--- program platizq (robot Fanuc LR Mate 200iD/7L) ---
  Suave(1)
  Establecer velocidad (1000.0 mm/s)
  Est. Ref.: RobotiQ 2F-140 Gripper (Mechanism) Base
  Est. herr: Tool 1
  Mostrar Tool 1
  MoveJ 1 to (260.93, 112.74, 317.18) mm, rotated rx -163.75 ry -45.95 rz -164.16 deg; joints [66.37, 34.682, -17.427, -50.975, -57.423, 69.366]
  MoveL 2 to (260.93, 112.74, 317.18) mm, rotated rx -163.75 ry -45.95 rz -164.16 deg; joints [66.37, 34.682, -17.427, -50.975, -57.423, 69.366]
  MoveL 3 to (241.32, 112.74, 219.12) mm, rotated rx -163.75 ry -45.95 rz -164.16 deg; joints [66.988, 41.165, -27.056, -56.554, -51.255, 78.508]
  MoveL 4 to (241.32, 112.74, 219.12) mm, rotated rx -163.75 ry -45.95 rz -164.16 deg; joints [66.988, 41.165, -27.056, -56.554, -51.255, 78.508]
  Establecer velocidad (50.0 mm/s)
  MoveL 5 to (253.05, 113.72, 219.12) mm, rotated rx -163.75 ry -45.95 rz -164.16 deg; joints [66.551, 39.855, -28.019, -57.172, -51.053, 79.816]
  MoveL 6 to (264.85, 113.71, 219.12) mm, rotated rx -163.75 ry -45.95 rz -164.16 deg; joints [66.172, 38.517, -28.983, -57.797, -50.815, 81.094]
  MoveL 7 to (276.61, 112.7, 219.12) mm, rotated rx -163.75 ry -45.95 rz -164.16 deg; joints [65.858, 37.162, -29.939, -58.425, -50.543, 82.329]
  MoveL 8 to (288.2, 110.7, 219.12) mm, rotated rx -163.75 ry -45.95 rz -164.16 deg; joints [65.614, 35.801, -30.876, -59.055, -50.236, 83.51]
  MoveL 9 to (299.55, 107.74, 219.66) mm, rotated rx -163.75 ry -45.95 rz -164.16 deg; joints [65.446, 34.407, -31.728, -59.642, -49.925, 84.562]
  MoveL 10 to (311.25, 103.8, 221.33) mm, rotated rx -163.75 ry -45.95 rz -164.16 deg; joints [65.334, 32.878, -32.469, -60.165, -49.635, 85.463]
  MoveL 11 to (322.85, 100.34, 224.12) mm, rotated rx -163.75 ry -45.95 rz -164.16 deg; joints [65.186, 31.325, -33.014, -60.541, -49.474, 86.167]
  MoveL 12 to (334.34, 97.51, 228.04) mm, rotated rx -163.75 ry -45.95 rz -164.16 deg; joints [64.983, 29.751, -33.357, -60.757, -49.454, 86.67]
  MoveL 13 to (346, 95.24, 231.53) mm, rotated rx -163.75 ry -45.95 rz -164.16 deg; joints [64.72, 28.217, -33.701, -60.96, -49.478, 87.205]
  MoveL 14 to (357.95, 93.53, 233.87) mm, rotated rx -163.75 ry -45.95 rz -164.16 deg; joints [64.39, 26.758, -34.143, -61.22, -49.504, 87.889]
  MoveL 15 to (370.19, 92.4, 235.02) mm, rotated rx -163.75 ry -45.95 rz -164.16 deg; joints [63.985, 25.377, -34.691, -61.538, -49.535, 88.731]
  MoveL 16 to (383.51, 91.88, 235.15) mm, rotated rx -163.75 ry -45.95 rz -164.16 deg; joints [63.465, 23.993, -35.369, -61.92, -49.589, 89.781]
  MoveL 17 to (396.84, 92.08, 235.15) mm, rotated rx -163.75 ry -45.95 rz -164.16 deg; joints [62.858, 22.663, -36.01, -62.244, -49.724, 90.827]
  MoveL 18 to (410.17, 92.08, 235.15) mm, rotated rx -163.75 ry -45.95 rz -164.16 deg; joints [62.245, 21.332, -36.621, -62.531, -49.879, 91.835]
  MoveL 19 to (423.5, 92.08, 235.15) mm, rotated rx -163.75 ry -45.95 rz -164.16 deg; joints [61.606, 20.009, -37.197, -62.774, -50.068, 92.81]
  MoveL 20 to (436.83, 92.08, 235.15) mm, rotated rx -163.75 ry -45.95 rz -164.16 deg; joints [60.939, 18.692, -37.738, -62.971, -50.292, 93.751]
  MoveL 21 to (445.16, 92.08, 235.15) mm, rotated rx -163.75 ry -45.95 rz -164.16 deg; joints [60.508, 17.872, -38.059, -63.071, -50.45, 94.323]
  MoveL 22 to (453.49, 92.08, 235.15) mm, rotated rx -163.75 ry -45.95 rz -164.16 deg; joints [60.065, 17.054, -38.366, -63.152, -50.622, 94.881]
  MoveL 23 to (461.82, 92.08, 235.15) mm, rotated rx -163.75 ry -45.95 rz -164.16 deg; joints [59.609, 16.238, -38.659, -63.214, -50.808, 95.427]
  MoveL 24 to (470.22, 91.84, 235.15) mm, rotated rx -163.75 ry -45.95 rz -164.16 deg; joints [59.16, 15.403, -38.947, -63.269, -50.991, 95.961]
  MoveL 25 to (476.05, 90.4, 235.15) mm, rotated rx -163.75 ry -45.95 rz -164.16 deg; joints [58.963, 14.749, -39.161, -63.356, -51.031, 96.296]
  MoveL 26 to (481.67, 87.57, 235.15) mm, rotated rx -163.75 ry -45.95 rz -164.16 deg; joints [58.91, 14.031, -39.387, -63.501, -50.967, 96.58]
  MoveL 27 to (486.6, 83.43, 235.15) mm, rotated rx -163.75 ry -45.95 rz -164.16 deg; joints [59.025, 13.302, -39.606, -63.701, -50.79, 96.782]
  MoveL 28 to (490.42, 78.28, 235.15) mm, rotated rx -163.75 ry -45.95 rz -164.16 deg; joints [59.311, 12.621, -39.801, -63.948, -50.507, 96.882]
  MoveL 29 to (492.88, 72.58, 235.15) mm, rotated rx -163.75 ry -45.95 rz -164.16 deg; joints [59.741, 12.041, -39.958, -64.221, -50.141, 96.879]
  MoveL 30 to (493.98, 66.8, 235.15) mm, rotated rx -163.75 ry -45.95 rz -164.16 deg; joints [60.268, 11.597, -40.075, -64.502, -49.727, 96.788]
  MoveL 31 to (494.07, 61.23, 235.15) mm, rotated rx -163.75 ry -45.95 rz -164.16 deg; joints [60.841, 11.27, -40.158, -64.774, -49.296, 96.64]
  MoveL 32 to (494.07, 55.68, 235.15) mm, rotated rx -163.75 ry -45.95 rz -164.16 deg; joints [61.423, 10.958, -40.235, -65.047, -48.86, 96.482]
  MoveL 33 to (493.53, 50, 235.15) mm, rotated rx -163.75 ry -45.95 rz -164.16 deg; joints [62.056, 10.7, -40.297, -65.328, -48.395, 96.287]
  MoveL 34 to (491.67, 44.21, 235.15) mm, rotated rx -163.75 ry -45.95 rz -164.16 deg; joints [62.78, 10.579, -40.325, -65.614, -47.881, 96.014]
  MoveL 35 to (488.43, 38.76, 235.15) mm, rotated rx -163.75 ry -45.95 rz -164.16 deg; joints [63.546, 10.629, -40.313, -65.88, -47.354, 95.675]
  MoveL 36 to (483.95, 34.13, 235.15) mm, rotated rx -163.75 ry -45.95 rz -164.16 deg; joints [64.285, 10.862, -40.258, -66.098, -46.861, 95.292]
  MoveL 37 to (478.57, 30.7, 235.15) mm, rotated rx -163.75 ry -45.95 rz -164.16 deg; joints [64.933, 11.256, -40.161, -66.244, -46.448, 94.895]
  MoveL 38 to (472.77, 28.65, 235.15) mm, rotated rx -163.75 ry -45.95 rz -164.16 deg; joints [65.443, 11.768, -40.03, -66.308, -46.143, 94.513]
  MoveL 39 to (465.18, 27.94, 235.15) mm, rotated rx -163.75 ry -45.95 rz -164.16 deg; joints [65.887, 12.534, -39.824, -66.279, -45.915, 94.061]
  MoveL 40 to (457.78, 27.94, 235.15) mm, rotated rx -163.75 ry -45.95 rz -164.16 deg; joints [66.235, 13.314, -39.602, -66.199, -45.759, 93.627]
  MoveL 41 to (450.37, 27.94, 235.15) mm, rotated rx -163.75 ry -45.95 rz -164.16 deg; joints [66.574, 14.092, -39.368, -66.103, -45.614, 93.18]
  MoveL 42 to (442.97, 27.94, 235.15) mm, rotated rx -163.75 ry -45.95 rz -164.16 deg; joints [66.905, 14.869, -39.122, -65.989, -45.48, 92.719]
  MoveL 43 to (435.56, 27.94, 235.15) mm, rotated rx -163.75 ry -45.95 rz -164.16 deg; joints [67.226, 15.646, -38.864, -65.859, -45.357, 92.245]
  MoveL 44 to (428.16, 27.94, 235.15) mm, rotated rx -163.75 ry -45.95 rz -164.16 deg; joints [67.539, 16.422, -38.594, -65.712, -45.245, 91.758]
  MoveL 45 to (413.49, 27.94, 235.15) mm, rotated rx -163.75 ry -45.95 rz -164.16 deg; joints [68.135, 17.958, -38.025, -65.374, -45.055, 90.755]
  MoveL 46 to (398.83, 27.94, 235.15) mm, rotated rx -163.75 ry -45.95 rz -164.16 deg; joints [68.702, 19.495, -37.412, -64.975, -44.906, 89.701]
  MoveL 47 to (384.18, 27.45, 235.15) mm, rotated rx -163.75 ry -45.95 rz -164.16 deg; joints [69.288, 21.014, -36.762, -64.536, -44.76, 88.584]
  MoveL 48 to (369.59, 25.97, 235) mm, rotated rx -163.75 ry -45.95 rz -164.16 deg; joints [69.936, 22.505, -36.108, -64.097, -44.573, 87.425]
  MoveL 49 to (357.46, 23.95, 233.79) mm, rotated rx -163.75 ry -45.95 rz -164.16 deg; joints [70.525, 23.796, -35.681, -63.837, -44.332, 86.577]
  MoveL 50 to (345.61, 21.29, 231.44) mm, rotated rx -163.75 ry -45.95 rz -164.16 deg; joints [71.143, 25.115, -35.39, -63.699, -44.01, 85.885]
  MoveL 51 to (334.07, 18.15, 227.95) mm, rotated rx -163.75 ry -45.95 rz -164.16 deg; joints [71.773, 26.466, -35.228, -63.675, -43.621, 85.346]
  MoveL 52 to (322.58, 15.47, 224.04) mm, rotated rx -163.75 ry -45.95 rz -164.16 deg; joints [72.34, 27.861, -35.073, -63.637, -43.274, 84.844]
  MoveL 53 to (310.79, 13.36, 221.24) mm, rotated rx -163.75 ry -45.95 rz -164.16 deg; joints [72.848, 29.241, -34.718, -63.39, -43.059, 84.107]
  MoveL 54 to (298.7, 11.85, 219.58) mm, rotated rx -163.75 ry -45.95 rz -164.16 deg; joints [73.295, 30.606, -34.158, -62.93, -42.983, 83.131]
  MoveL 55 to (287.65, 11.04, 219.12) mm, rotated rx -163.75 ry -45.95 rz -164.16 deg; joints [73.643, 31.816, -33.482, -62.337, -43.037, 82.057]
  MoveL 56 to (276.52, 10.76, 219.12) mm, rotated rx -163.75 ry -45.95 rz -164.16 deg; joints [73.937, 33.036, -32.706, -61.643, -43.184, 80.886]
  MoveL 57 to (265.38, 10.76, 219.12) mm, rotated rx -163.75 ry -45.95 rz -164.16 deg; joints [74.199, 34.28, -31.895, -60.914, -43.38, 79.692]
  MoveL 58 to (254.26, 11.36, 219.12) mm, rotated rx -163.75 ry -45.95 rz -164.16 deg; joints [74.404, 35.558, -31.04, -60.146, -43.648, 78.486]
  MoveL 59 to (243.27, 13.24, 219.12) mm, rotated rx -163.75 ry -45.95 rz -164.16 deg; joints [74.498, 36.878, -30.135, -59.338, -44.034, 77.299]
  MoveL 60 to (232.6, 16.36, 219.32) mm, rotated rx -163.75 ry -45.95 rz -164.16 deg; joints [74.486, 38.214, -29.168, -58.488, -44.543, 76.121]
  MoveL 61 to (222.4, 20.67, 219.99) mm, rotated rx -163.75 ry -45.95 rz -164.16 deg; joints [74.372, 39.53, -28.125, -57.598, -45.18, 74.941]
  MoveL 62 to (212.73, 26.14, 221.07) mm, rotated rx -163.75 ry -45.95 rz -164.16 deg; joints [74.162, 40.83, -27.015, -56.685, -45.938, 73.777]
  MoveL 63 to (203.82, 32.62, 222.45) mm, rotated rx -163.75 ry -45.95 rz -164.16 deg; joints [73.867, 42.091, -25.876, -55.791, -46.791, 72.672]
  MoveL 64 to (198.88, 36.96, 223.38) mm, rotated rx -163.75 ry -45.95 rz -164.16 deg; joints [73.652, 42.825, -25.188, -55.273, -47.34, 72.046]
  MoveL 65 to (194.23, 41.63, 224.35) mm, rotated rx -163.75 ry -45.95 rz -164.16 deg; joints [73.409, 43.547, -24.498, -54.77, -47.917, 71.452]
  MoveL 66 to (189.92, 46.67, 225.35) mm, rotated rx -163.75 ry -45.95 rz -164.16 deg; joints [73.136, 44.252, -23.813, -54.289, -48.517, 70.898]
  MoveL 67 to (186.72, 52.48, 226.16) mm, rotated rx -163.75 ry -45.95 rz -164.16 deg; joints [72.787, 44.867, -23.221, -53.895, -49.123, 70.51]
  MoveL 68 to (185.04, 58.92, 226.6) mm, rotated rx -163.75 ry -45.95 rz -164.16 deg; joints [72.362, 45.336, -22.794, -53.631, -49.691, 70.36]
  MoveL 69 to (184.83, 66.37, 226.66) mm, rotated rx -163.75 ry -45.95 rz -164.16 deg; joints [71.836, 45.682, -22.514, -53.482, -50.247, 70.444]
  MoveL 70 to (185.41, 73.79, 226.5) mm, rotated rx -163.75 ry -45.95 rz -164.16 deg; joints [71.297, 45.942, -22.332, -53.401, -50.756, 70.64]
  MoveL 71 to (187.29, 80.95, 226.01) mm, rotated rx -163.75 ry -45.95 rz -164.16 deg; joints [70.746, 46.04, -22.325, -53.433, -51.17, 71.023]
  MoveL 72 to (190.4, 87.61, 225.24) mm, rotated rx -163.75 ry -45.95 rz -164.16 deg; joints [70.2, 45.976, -22.486, -53.568, -51.48, 71.573]
  MoveL 73 to (194.64, 93.62, 224.26) mm, rotated rx -163.75 ry -45.95 rz -164.16 deg; joints [69.67, 45.75, -22.802, -53.797, -51.687, 72.268]
  MoveL 74 to (199.85, 98.76, 223.19) mm, rotated rx -163.75 ry -45.95 rz -164.16 deg; joints [69.172, 45.372, -23.254, -54.102, -51.792, 73.077]
  MoveL 75 to (205.9, 102.91, 222.1) mm, rotated rx -163.75 ry -45.95 rz -164.16 deg; joints [68.717, 44.852, -23.817, -54.472, -51.802, 73.968]
  MoveL 76 to (212.58, 105.92, 221.09) mm, rotated rx -163.75 ry -45.95 rz -164.16 deg; joints [68.319, 44.205, -24.463, -54.89, -51.724, 74.907]
  MoveL 77 to (219.61, 108.2, 220.26) mm, rotated rx -163.75 ry -45.95 rz -164.16 deg; joints [67.958, 43.487, -25.137, -55.324, -51.608, 75.85]
  MoveL 78 to (226.74, 110.09, 219.65) mm, rotated rx -163.75 ry -45.95 rz -164.16 deg; joints [67.616, 42.741, -25.794, -55.746, -51.49, 76.765]
  MoveL 79 to (233.98, 111.61, 219.26) mm, rotated rx -163.75 ry -45.95 rz -164.16 deg; joints [67.293, 41.968, -26.434, -56.156, -51.373, 77.652]
  MoveL 80 to (241.32, 112.74, 219.12) mm, rotated rx -163.75 ry -45.95 rz -164.16 deg; joints [66.988, 41.165, -27.056, -56.554, -51.255, 78.508]
  Establecer velocidad (1000.0 mm/s)
  MoveL 81 to (241.32, 112.74, 219.12) mm, rotated rx -163.75 ry -45.95 rz -164.16 deg; joints [66.988, 41.165, -27.056, -56.554, -51.255, 78.508]
  MoveL 82 to (260.93, 112.74, 317.18) mm, rotated rx -163.75 ry -45.95 rz -164.16 deg; joints [66.37, 34.682, -17.427, -50.975, -57.423, 69.366]
  Establecer velocidad (1000.0 mm/s)
  MoveL 83 to (452.25, 27.76, 382.46) mm, rotated rx -163.75 ry -45.95 rz -164.16 deg; joints [66.508, 5.685, -18.926, -51.728, -56.385, 70.666]
  MoveL 84 to (432.64, 27.76, 284.4) mm, rotated rx -163.75 ry -45.95 rz -164.16 deg; joints [67.369, 12.539, -31.994, -60.148, -48.379, 83.782]
  MoveL 85 to (432.64, 27.76, 284.4) mm, rotated rx -163.75 ry -45.95 rz -164.16 deg; joints [67.369, 12.539, -31.994, -60.148, -48.379, 83.782]
  Establecer velocidad (50.0 mm/s)
  MoveL 86 to (452.8, 28.72, 284.4) mm, rotated rx -163.75 ry -45.95 rz -164.16 deg; joints [66.383, 10.356, -32.504, -60.376, -48.85, 84.924]
  MoveL 87 to (472.8, 31.52, 284.4) mm, rotated rx -163.75 ry -45.95 rz -164.16 deg; joints [65.133, 8.281, -32.901, -60.447, -49.569, 86.066]
  MoveL 88 to (479.3, 33.32, 284.4) mm, rotated rx -163.75 ry -45.95 rz -164.16 deg; joints [64.612, 7.655, -33.003, -60.422, -49.899, 86.466]
  MoveL 89 to (485.2, 36.51, 284.4) mm, rotated rx -163.75 ry -45.95 rz -164.16 deg; joints [63.96, 7.172, -33.077, -60.346, -50.337, 86.901]
  MoveL 90 to (490.31, 40.91, 284.4) mm, rotated rx -163.75 ry -45.95 rz -164.16 deg; joints [63.21, 6.849, -33.124, -60.226, -50.859, 87.357]
  MoveL 91 to (494.31, 46.34, 284.4) mm, rotated rx -163.75 ry -45.95 rz -164.16 deg; joints [62.404, 6.717, -33.143, -60.069, -51.436, 87.809]
  MoveL 92 to (496.77, 52.59, 284.4) mm, rotated rx -163.75 ry -45.95 rz -164.16 deg; joints [61.595, 6.811, -33.13, -59.885, -52.029, 88.226]
  MoveL 93 to (497.4, 59.25, 284.4) mm, rotated rx -163.75 ry -45.95 rz -164.16 deg; joints [60.853, 7.137, -33.083, -59.69, -52.589, 88.57]
  MoveL 94 to (497.21, 64.6, 284.4) mm, rotated rx -163.75 ry -45.95 rz -164.16 deg; joints [60.305, 7.479, -33.031, -59.534, -53.012, 88.806]
  MoveL 95 to (495.99, 69.73, 284.4) mm, rotated rx -163.75 ry -45.95 rz -164.16 deg; joints [59.846, 7.923, -32.961, -59.385, -53.379, 88.975]
  MoveL 96 to (493.74, 74.55, 284.4) mm, rotated rx -163.75 ry -45.95 rz -164.16 deg; joints [59.489, 8.458, -32.871, -59.247, -53.683, 89.068]
  MoveL 97 to (490.6, 78.79, 284.4) mm, rotated rx -163.75 ry -45.95 rz -164.16 deg; joints [59.249, 9.05, -32.764, -59.125, -53.911, 89.083]
  MoveL 98 to (486.76, 82.45, 284.4) mm, rotated rx -163.75 ry -45.95 rz -164.16 deg; joints [59.112, 9.678, -32.643, -59.019, -54.071, 89.028]
  MoveL 99 to (480.86, 86.17, 284.4) mm, rotated rx -163.75 ry -45.95 rz -164.16 deg; joints [59.093, 10.521, -32.469, -58.907, -54.175, 88.854]
  MoveL 100 to (474.22, 88.37, 284.4) mm, rotated rx -163.75 ry -45.95 rz -164.16 deg; joints [59.264, 11.343, -32.285, -58.831, -54.146, 88.568]
  MoveL 101 to (467.32, 89.52, 284.4) mm, rotated rx -163.75 ry -45.95 rz -164.16 deg; joints [59.546, 12.127, -32.098, -58.775, -54.04, 88.218]
  MoveL 102 to (460.39, 90.46, 284.4) mm, rotated rx -163.75 ry -45.95 rz -164.16 deg; joints [59.842, 12.9, -31.901, -58.715, -53.927, 87.849]
  MoveL 103 to (453.43, 91.18, 284.4) mm, rotated rx -163.75 ry -45.95 rz -164.16 deg; joints [60.152, 13.663, -31.696, -58.651, -53.808, 87.462]
  MoveL 104 to (446.45, 91.7, 284.4) mm, rotated rx -163.75 ry -45.95 rz -164.16 deg; joints [60.476, 14.416, -31.482, -58.581, -53.685, 87.058]
  MoveL 105 to (429.96, 92.12, 284.4) mm, rotated rx -163.75 ry -45.95 rz -164.16 deg; joints [61.282, 16.152, -30.948, -58.396, -53.375, 86.043]
  MoveL 106 to (413.48, 91.53, 284.4) mm, rotated rx -163.75 ry -45.95 rz -164.16 deg; joints [62.137, 17.84, -30.376, -58.179, -53.05, 84.952]
  MoveL 107 to (403.76, 90.49, 284.4) mm, rotated rx -163.75 ry -45.95 rz -164.16 deg; joints [62.684, 18.804, -30.026, -58.041, -52.834, 84.267]
  MoveL 108 to (394.19, 88.84, 284.4) mm, rotated rx -163.75 ry -45.95 rz -164.16 deg; joints [63.262, 19.726, -29.675, -57.9, -52.595, 83.559]
  MoveL 109 to (384.65, 87.33, 284.4) mm, rotated rx -163.75 ry -45.95 rz -164.16 deg; joints [63.811, 20.66, -29.304, -57.734, -52.389, 82.843]
  MoveL 110 to (374.95, 87.44, 284.4) mm, rotated rx -163.75 ry -45.95 rz -164.16 deg; joints [64.212, 21.702, -28.873, -57.503, -52.323, 82.146]
  MoveL 111 to (365.25, 87.59, 284.4) mm, rotated rx -163.75 ry -45.95 rz -164.16 deg; joints [64.598, 22.751, -28.42, -57.252, -52.282, 81.433]
  MoveL 112 to (355.55, 87.57, 284.4) mm, rotated rx -163.75 ry -45.95 rz -164.16 deg; joints [64.987, 23.799, -27.949, -56.986, -52.25, 80.697]
  MoveL 113 to (351.15, 87.43, 284.4) mm, rotated rx -163.75 ry -45.95 rz -164.16 deg; joints [65.171, 24.271, -27.731, -56.861, -52.233, 80.354]
  MoveL 114 to (346.75, 87.18, 284.4) mm, rotated rx -163.75 ry -45.95 rz -164.16 deg; joints [65.362, 24.738, -27.511, -56.736, -52.211, 80.004]
  MoveL 115 to (342.36, 86.74, 284.4) mm, rotated rx -163.75 ry -45.95 rz -164.16 deg; joints [65.565, 25.196, -27.293, -56.611, -52.181, 79.647]
  MoveL 116 to (338.08, 85.69, 284.4) mm, rotated rx -163.75 ry -45.95 rz -164.16 deg; joints [65.813, 25.614, -27.09, -56.498, -52.108, 79.28]
  MoveL 117 to (334.49, 83.14, 284.4) mm, rotated rx -163.75 ry -45.95 rz -164.16 deg; joints [66.158, 25.885, -26.957, -56.436, -51.926, 78.924]
  MoveL 118 to (332.28, 80.19, 284.4) mm, rotated rx -163.75 ry -45.95 rz -164.16 deg; joints [66.483, 25.986, -26.907, -56.424, -51.712, 78.667]
  MoveL 119 to (331.08, 76.71, 284.4) mm, rotated rx -163.75 ry -45.95 rz -164.16 deg; joints [66.815, 25.953, -26.924, -56.456, -51.456, 78.475]
  MoveL 120 to (331.16, 73.04, 284.4) mm, rotated rx -163.75 ry -45.95 rz -164.16 deg; joints [67.118, 25.771, -27.013, -56.534, -51.181, 78.38]
  MoveL 121 to (332.81, 67.76, 284.4) mm, rotated rx -163.75 ry -45.95 rz -164.16 deg; joints [67.503, 25.341, -27.222, -56.698, -50.78, 78.362]
  MoveL 122 to (334.61, 62.54, 284.4) mm, rotated rx -163.75 ry -45.95 rz -164.16 deg; joints [67.883, 24.902, -27.433, -56.865, -50.382, 78.351]
  MoveL 123 to (334.06, 60.19, 284.4) mm, rotated rx -163.75 ry -45.95 rz -164.16 deg; joints [68.102, 24.858, -27.454, -56.892, -50.208, 78.236]
  MoveL 124 to (333.37, 57.83, 284.4) mm, rotated rx -163.75 ry -45.95 rz -164.16 deg; joints [68.327, 24.83, -27.467, -56.914, -50.034, 78.109]
  MoveL 125 to (332.69, 55.47, 284.4) mm, rotated rx -163.75 ry -45.95 rz -164.16 deg; joints [68.552, 24.802, -27.481, -56.936, -49.859, 77.981]
  MoveL 126 to (332.02, 53.1, 284.4) mm, rotated rx -163.75 ry -45.95 rz -164.16 deg; joints [68.776, 24.773, -27.494, -56.957, -49.685, 77.853]
  MoveL 127 to (331.37, 50.73, 284.4) mm, rotated rx -163.75 ry -45.95 rz -164.16 deg; joints [69.001, 24.743, -27.508, -56.979, -49.51, 77.726]
  MoveL 128 to (330.99, 48.32, 284.4) mm, rotated rx -163.75 ry -45.95 rz -164.16 deg; joints [69.221, 24.682, -27.537, -57.01, -49.331, 77.618]
  MoveL 129 to (331.56, 43.51, 284.4) mm, rotated rx -163.75 ry -45.95 rz -164.16 deg; joints [69.618, 24.415, -27.663, -57.12, -48.967, 77.505]
  MoveL 130 to (333.68, 39.14, 284.4) mm, rotated rx -163.75 ry -45.95 rz -164.16 deg; joints [69.931, 23.996, -27.858, -57.278, -48.629, 77.523]
  MoveL 131 to (336.88, 35.49, 284.4) mm, rotated rx -163.75 ry -45.95 rz -164.16 deg; joints [70.148, 23.487, -28.091, -57.461, -48.342, 77.647]
  MoveL 132 to (341.1, 33.11, 284.4) mm, rotated rx -163.75 ry -45.95 rz -164.16 deg; joints [70.224, 22.917, -28.346, -57.658, -48.148, 77.888]
  MoveL 133 to (345.9, 32.32, 284.4) mm, rotated rx -163.75 ry -45.95 rz -164.16 deg; joints [70.141, 22.346, -28.597, -57.843, -48.076, 78.224]
  MoveL 134 to (350.74, 31.87, 284.4) mm, rotated rx -163.75 ry -45.95 rz -164.16 deg; joints [70.024, 21.785, -28.837, -58.019, -48.036, 78.572]
  MoveL 135 to (355.61, 31.66, 284.4) mm, rotated rx -163.75 ry -45.95 rz -164.16 deg; joints [69.883, 21.233, -29.069, -58.186, -48.018, 78.924]
  MoveL 136 to (360.47, 31.61, 284.4) mm, rotated rx -163.75 ry -45.95 rz -164.16 deg; joints [69.725, 20.689, -29.292, -58.346, -48.018, 79.277]
  MoveL 137 to (365.34, 31.66, 284.4) mm, rotated rx -163.75 ry -45.95 rz -164.16 deg; joints [69.554, 20.149, -29.508, -58.498, -48.031, 79.63]
  MoveL 138 to (370.79, 31.8, 284.4) mm, rotated rx -163.75 ry -45.95 rz -164.16 deg; joints [69.353, 19.55, -29.743, -58.66, -48.059, 80.021]
  MoveL 139 to (376.24, 31.99, 284.4) mm, rotated rx -163.75 ry -45.95 rz -164.16 deg; joints [69.144, 18.953, -29.969, -58.814, -48.096, 80.408]
  MoveL 140 to (381.69, 32.16, 284.4) mm, rotated rx -163.75 ry -45.95 rz -164.16 deg; joints [68.933, 18.357, -30.189, -58.962, -48.139, 80.788]
  MoveL 141 to (387.14, 32.28, 284.4) mm, rotated rx -163.75 ry -45.95 rz -164.16 deg; joints [68.722, 17.76, -30.404, -59.104, -48.184, 81.16]
  MoveL 142 to (392.5, 31.25, 284.4) mm, rotated rx -163.75 ry -45.95 rz -164.16 deg; joints [68.622, 17.124, -30.624, -59.262, -48.145, 81.474]
  MoveL 143 to (397.9, 29.94, 284.4) mm, rotated rx -163.75 ry -45.95 rz -164.16 deg; joints [68.544, 16.472, -30.844, -59.422, -48.091, 81.773]
  MoveL 144 to (403.83, 28.61, 284.4) mm, rotated rx -163.75 ry -45.95 rz -164.16 deg; joints [68.447, 15.758, -31.074, -59.589, -48.046, 82.097]
  MoveL 145 to (408.55, 28, 284.4) mm, rotated rx -163.75 ry -45.95 rz -164.16 deg; joints [68.324, 15.211, -31.244, -59.705, -48.051, 82.366]
  MoveL 146 to (412.24, 27.79, 284.4) mm, rotated rx -163.75 ry -45.95 rz -164.16 deg; joints [68.2, 14.793, -31.37, -59.786, -48.079, 82.584]
  MoveL 147 to (415.69, 27.76, 284.4) mm, rotated rx -163.75 ry -45.95 rz -164.16 deg; joints [68.066, 14.411, -31.483, -59.855, -48.121, 82.792]
  MoveL 148 to (418.69, 27.76, 284.4) mm, rotated rx -163.75 ry -45.95 rz -164.16 deg; joints [67.946, 14.08, -31.578, -59.912, -48.162, 82.971]
  MoveL 149 to (422.53, 27.76, 284.4) mm, rotated rx -163.75 ry -45.95 rz -164.16 deg; joints [67.79, 13.656, -31.697, -59.982, -48.217, 83.199]
  MoveL 150 to (427.35, 27.76, 284.4) mm, rotated rx -163.75 ry -45.95 rz -164.16 deg; joints [67.591, 13.123, -31.842, -60.064, -48.292, 83.48]
  MoveL 151 to (432.64, 27.76, 284.4) mm, rotated rx -163.75 ry -45.95 rz -164.16 deg; joints [67.369, 12.539, -31.994, -60.148, -48.379, 83.782]
  Establecer velocidad (1000.0 mm/s)
  MoveL 152 to (432.64, 27.76, 284.4) mm, rotated rx -163.75 ry -45.95 rz -164.16 deg; joints [67.369, 12.539, -31.994, -60.148, -48.379, 83.782]
  MoveL 153 to (452.25, 27.76, 382.46) mm, rotated rx -163.75 ry -45.95 rz -164.16 deg; joints [66.508, 5.685, -18.926, -51.728, -56.385, 70.666]

--- program carribizq (robot Fanuc LR Mate 200iD/7L) ---
  Suave(1)
  Establecer velocidad (1000.0 mm/s)
  Est. Ref.: RobotiQ 2F-140 Gripper (Mechanism) Base
  Est. herr: Tool 1
  Mostrar Tool 1
  MoveJ 1 to (259.22, -163.5, 158.15) mm, rotated rx 167 ry 29.36 rz -96.45 deg; joints [108.037, 52.448, -19.707, 33.515, -72.983, 58.084]
  MoveL 2 to (259.22, -163.5, 158.15) mm, rotated rx 167 ry 29.36 rz -96.45 deg; joints [108.037, 52.448, -19.707, 33.515, -72.983, 58.084]
  MoveL 3 to (239.61, -163.5, 60.09) mm, rotated rx 167 ry 29.36 rz -96.45 deg; joints [107.615, 60.488, -26.388, 34.925, -67.238, 54.431]
  MoveL 4 to (239.61, -163.5, 60.09) mm, rotated rx 167 ry 29.36 rz -96.45 deg; joints [107.615, 60.488, -26.388, 34.925, -67.238, 54.431]
  Establecer velocidad (50.0 mm/s)
  MoveL 5 to (229.89, -163.5, 58.94) mm, rotated rx 167 ry 29.36 rz -96.45 deg; joints [107.413, 62.037, -25.037, 34.636, -68.244, 55.425]
  MoveL 6 to (220.16, -163.5, 57.58) mm, rotated rx 167 ry 29.36 rz -96.45 deg; joints [107.215, 63.684, -23.61, 34.346, -69.318, 56.452]
  MoveL 7 to (209.4, -163.5, 55.83) mm, rotated rx 167 ry 29.36 rz -96.45 deg; joints [107.001, 65.643, -21.916, 34.023, -70.608, 57.638]
  MoveL 8 to (197.24, -163.5, 53.55) mm, rotated rx 167 ry 29.36 rz -96.45 deg; joints [106.766, 68.074, -19.81, 33.651, -72.235, 59.068]
  MoveL 9 to (186.82, -163.5, 51.32) mm, rotated rx 167 ry 29.36 rz -96.45 deg; joints [106.569, 70.407, -17.775, 33.324, -73.829, 60.405]
  MoveL 10 to (181.89, -163.5, 50.18) mm, rotated rx 167 ry 29.36 rz -96.45 deg; joints [106.477, 71.62, -16.708, 33.166, -74.674, 61.089]
  MoveL 11 to (177.52, -163.5, 49.12) mm, rotated rx 167 ry 29.36 rz -96.45 deg; joints [106.397, 72.773, -15.685, 33.022, -75.489, 61.733]
  MoveL 12 to (175.68, -163.5, 48.58) mm, rotated rx 167 ry 29.36 rz -96.45 deg; joints [106.363, 73.287, -15.237, 32.962, -75.847, 62.013]
  MoveL 13 to (174.49, -163.5, 47.81) mm, rotated rx 167 ry 29.36 rz -96.45 deg; joints [106.341, 73.65, -14.975, 32.927, -76.055, 62.178]
  MoveL 14 to (173.49, -163.5, 46.5) mm, rotated rx 167 ry 29.36 rz -96.45 deg; joints [106.323, 73.997, -14.803, 32.905, -76.19, 62.29]
  MoveL 15 to (173.06, -163.5, 45.24) mm, rotated rx 167 ry 29.36 rz -96.45 deg; joints [106.315, 74.182, -14.787, 32.904, -76.2, 62.305]
  MoveL 16 to (172.98, -163.5, 43.71) mm, rotated rx 167 ry 29.36 rz -96.45 deg; joints [106.314, 74.283, -14.895, 32.918, -76.109, 62.246]
  MoveL 17 to (172.98, -163.5, 41.64) mm, rotated rx 167 ry 29.36 rz -96.45 deg; joints [106.314, 74.393, -15.069, 32.942, -75.963, 62.149]
  MoveL 18 to (172.98, -163.5, 37.97) mm, rotated rx 167 ry 29.36 rz -96.45 deg; joints [106.314, 74.591, -15.374, 32.984, -75.707, 61.978]
  MoveL 19 to (172.98, -163.5, 33.71) mm, rotated rx 167 ry 29.36 rz -96.45 deg; joints [106.314, 74.828, -15.721, 33.032, -75.415, 61.782]
  MoveL 20 to (172.98, -163.5, 29.44) mm, rotated rx 167 ry 29.36 rz -96.45 deg; joints [106.314, 75.071, -16.063, 33.081, -75.129, 61.59]
  MoveL 21 to (172.98, -163.5, 25.06) mm, rotated rx 167 ry 29.36 rz -96.45 deg; joints [106.314, 75.327, -16.406, 33.132, -74.841, 61.395]
  Establecer velocidad (1000.0 mm/s)
  MoveL 22 to (172.98, -163.5, 25.06) mm, rotated rx 167 ry 29.36 rz -96.45 deg; joints [106.314, 75.327, -16.406, 33.132, -74.841, 61.395]
  MoveL 23 to (192.59, -163.5, 123.12) mm, rotated rx 167 ry 29.36 rz -96.45 deg; joints [106.677, 65.939, -12.253, 32.578, -78.522, 63.407]
  Establecer velocidad (1000.0 mm/s)
  MoveL 24 to (269.02, -163.5, 159.11) mm, rotated rx 167 ry 29.36 rz -96.45 deg; joints [108.255, 50.959, -20.839, 33.69, -72.153, 57.248]
  MoveL 25 to (249.41, -163.5, 61.05) mm, rotated rx 167 ry 29.36 rz -96.45 deg; joints [107.824, 59.011, -27.687, 35.216, -66.282, 53.453]
  MoveL 26 to (249.41, -163.5, 61.05) mm, rotated rx 167 ry 29.36 rz -96.45 deg; joints [107.824, 59.011, -27.687, 35.216, -66.282, 53.453]
  Establecer velocidad (50.0 mm/s)
  MoveL 27 to (267.91, -163.5, 63.56) mm, rotated rx 167 ry 29.36 rz -96.45 deg; joints [108.231, 56.337, -29.895, 35.737, -64.69, 51.726]
  MoveL 28 to (288.24, -163.5, 68.51) mm, rotated rx 167 ry 29.36 rz -96.45 deg; joints [108.699, 53.442, -31.899, 36.23, -63.305, 50.054]
  MoveL 29 to (307.9, -163.5, 75.65) mm, rotated rx 167 ry 29.36 rz -96.45 deg; joints [109.174, 50.62, -33.429, 36.605, -62.311, 48.671]
  MoveL 30 to (326.67, -163.5, 84.9) mm, rotated rx 167 ry 29.36 rz -96.45 deg; joints [109.65, 47.853, -34.495, 36.847, -61.693, 47.59]
  MoveL 31 to (344.31, -163.5, 96.14) mm, rotated rx 167 ry 29.36 rz -96.45 deg; joints [110.119, 45.139, -35.104, 36.944, -61.437, 46.824]
  MoveL 32 to (360.62, -163.5, 109.24) mm, rotated rx 167 ry 29.36 rz -96.45 deg; joints [110.572, 42.486, -35.262, 36.895, -61.532, 46.38]
  MoveL 33 to (375.4, -163.5, 124.04) mm, rotated rx 167 ry 29.36 rz -96.45 deg; joints [110.999, 39.913, -34.98, 36.709, -61.968, 46.254]
  Establecer velocidad (1000.0 mm/s)
  MoveL 34 to (375.4, -163.5, 124.04) mm, rotated rx 167 ry 29.36 rz -96.45 deg; joints [110.999, 39.913, -34.98, 36.709, -61.968, 46.254]
  MoveL 35 to (395.01, -163.5, 222.1) mm, rotated rx 167 ry 29.36 rz -96.45 deg; joints [111.592, 32.136, -25.489, 34.139, -70.007, 51.814]
  Establecer velocidad (1000.0 mm/s)
  MoveL 36 to (503.79, -163.5, 187.74) mm, rotated rx 167 ry 29.36 rz -96.45 deg; joints [115.563, 22.393, -35.87, 35.881, -63.453, 42.289]
  MoveL 37 to (484.18, -163.5, 89.68) mm, rotated rx 167 ry 29.36 rz -96.45 deg; joints [114.75, 31.996, -46.786, 40.191, -54.465, 35.007]
  MoveL 38 to (484.18, -163.5, 89.68) mm, rotated rx 167 ry 29.36 rz -96.45 deg; joints [114.75, 31.996, -46.786, 40.191, -54.465, 35.007]
  Establecer velocidad (50.0 mm/s)
  MoveL 39 to (486.5, -163.5, 73.75) mm, rotated rx 167 ry 29.36 rz -96.45 deg; joints [114.843, 33.232, -48.798, 41.119, -52.979, 33.322]
  MoveL 40 to (486.54, -163.5, 57.65) mm, rotated rx 167 ry 29.36 rz -96.45 deg; joints [114.845, 34.738, -50.649, 42.068, -51.595, 31.768]
  MoveL 41 to (484.29, -163.5, 41.71) mm, rotated rx 167 ry 29.36 rz -96.45 deg; joints [114.754, 36.463, -52.281, 42.999, -50.355, 30.402]
  MoveL 42 to (482.22, -163.5, 33.56) mm, rotated rx 167 ry 29.36 rz -96.45 deg; joints [114.671, 37.432, -53.026, 43.462, -49.777, 29.783]
  Establecer velocidad (1000.0 mm/s)
  MoveL 43 to (482.22, -163.5, 33.56) mm, rotated rx 167 ry 29.36 rz -96.45 deg; joints [114.671, 37.432, -53.026, 43.462, -49.777, 29.783]
  MoveL 44 to (501.83, -163.5, 131.62) mm, rotated rx 167 ry 29.36 rz -96.45 deg; joints [115.479, 26.799, -42.817, 38.262, -57.868, 37.546]
  Establecer velocidad (1000.0 mm/s)
  MoveL 45 to (503.79, -163.5, 187.74) mm, rotated rx 167 ry 29.36 rz -96.45 deg; joints [115.563, 22.393, -35.87, 35.881, -63.453, 42.289]
  MoveL 46 to (484.18, -163.5, 89.68) mm, rotated rx 167 ry 29.36 rz -96.45 deg; joints [114.75, 31.996, -46.786, 40.191, -54.465, 35.007]
  MoveL 47 to (484.18, -163.5, 89.68) mm, rotated rx 167 ry 29.36 rz -96.45 deg; joints [114.75, 31.996, -46.786, 40.191, -54.465, 35.007]
  Establecer velocidad (50.0 mm/s)
  MoveL 48 to (477.64, -163.5, 124.04) mm, rotated rx 167 ry 29.36 rz -96.45 deg; joints [114.489, 29.7, -42.306, 38.373, -57.816, 38.596]
  Establecer velocidad (1000.0 mm/s)
  MoveL 49 to (477.64, -163.5, 124.04) mm, rotated rx 167 ry 29.36 rz -96.45 deg; joints [114.489, 29.7, -42.306, 38.373, -57.816, 38.596]
  MoveL 50 to (497.25, -163.5, 222.1) mm, rotated rx 167 ry 29.36 rz -96.45 deg; joints [115.286, 20.903, -31.195, 34.704, -67.136, 45.469]

--- program cerlatder (robot Fanuc LR Mate 200iD/7L) ---
  Suave(1)
  Establecer velocidad (1000.0 mm/s)
  Est. Ref.: RobotiQ 2F-140 Gripper (Mechanism) Base
  Est. herr: Tool 1
  Mostrar Tool 1
  MoveJ 1 to (288.05, 234.2, 246.85) mm, rotated rx 165.67 ry -43.82 rz -104.8 deg; joints [59.121, 45.327, -18.732, -47.862, -74.104, 115.327]
  MoveL 2 to (288.05, 234.2, 246.85) mm, rotated rx 165.67 ry -43.82 rz -104.8 deg; joints [59.121, 45.327, -18.732, -47.862, -74.104, 115.327]
  MoveL 3 to (268.44, 234.2, 148.79) mm, rotated rx 165.67 ry -43.82 rz -104.8 deg; joints [59.852, 52.376, -26.936, -50.112, -68.205, 121.398]
  MoveL 4 to (268.44, 234.2, 148.79) mm, rotated rx 165.67 ry -43.82 rz -104.8 deg; joints [59.852, 52.376, -26.936, -50.112, -68.205, 121.398]
  Establecer velocidad (50.0 mm/s)
  MoveL 5 to (280.02, 235.56, 148.79) mm, rotated rx 165.67 ry -43.82 rz -104.8 deg; joints [59.338, 51.098, -28.072, -50.345, -67.829, 122.654]
  MoveL 6 to (291.68, 235.7, 148.79) mm, rotated rx 165.67 ry -43.82 rz -104.8 deg; joints [58.886, 49.776, -29.235, -50.602, -67.394, 123.897]
  MoveL 7 to (303.33, 235.61, 148.79) mm, rotated rx 165.67 ry -43.82 rz -104.8 deg; joints [58.438, 48.483, -30.362, -50.85, -66.982, 125.111]
  MoveL 8 to (314.96, 234.96, 148.99) mm, rotated rx 165.67 ry -43.82 rz -104.8 deg; joints [58.015, 47.185, -31.451, -51.093, -66.578, 126.28]
  MoveL 9 to (327.03, 233.66, 150.27) mm, rotated rx 165.67 ry -43.82 rz -104.8 deg; joints [57.605, 45.765, -32.464, -51.316, -66.215, 127.379]
  MoveL 10 to (338.81, 231.75, 152.7) mm, rotated rx 165.67 ry -43.82 rz -104.8 deg; joints [57.235, 44.294, -33.32, -51.499, -65.923, 128.324]
  MoveL 11 to (350.29, 229.26, 156.27) mm, rotated rx 165.67 ry -43.82 rz -104.8 deg; joints [56.906, 42.767, -34.02, -51.639, -65.703, 129.112]
  MoveL 12 to (361.65, 226.21, 160.06) mm, rotated rx 165.67 ry -43.82 rz -104.8 deg; joints [56.609, 41.221, -34.669, -51.772, -65.493, 129.837]
  MoveL 13 to (373.3, 223.38, 162.74) mm, rotated rx 165.67 ry -43.82 rz -104.8 deg; joints [56.275, 39.755, -35.399, -51.92, -65.257, 130.655]
  MoveL 14 to (385.24, 221.18, 164.28) mm, rotated rx 165.67 ry -43.82 rz -104.8 deg; joints [55.872, 38.395, -36.198, -52.07, -65.023, 131.57]
  MoveL 15 to (398.34, 219.58, 164.67) mm, rotated rx 165.67 ry -43.82 rz -104.8 deg; joints [55.359, 37.067, -37.136, -52.228, -64.772, 132.667]
  MoveL 16 to (411.52, 218.78, 164.67) mm, rotated rx 165.67 ry -43.82 rz -104.8 deg; joints [54.765, 35.831, -38.048, -52.343, -64.587, 133.783]
  MoveL 17 to (424.74, 218.69, 164.67) mm, rotated rx 165.67 ry -43.82 rz -104.8 deg; joints [54.099, 34.661, -38.895, -52.4, -64.483, 134.88]
  MoveL 18 to (437.95, 218.69, 164.67) mm, rotated rx 165.67 ry -43.82 rz -104.8 deg; joints [53.404, 33.518, -39.707, -52.424, -64.413, 135.956]
  MoveL 19 to (451.16, 218.69, 164.67) mm, rotated rx 165.67 ry -43.82 rz -104.8 deg; joints [52.685, 32.395, -40.489, -52.419, -64.372, 137.015]
  MoveL 20 to (484.19, 218.69, 164.67) mm, rotated rx 165.67 ry -43.82 rz -104.8 deg; joints [50.779, 29.672, -42.315, -52.271, -64.388, 139.587]
  MoveL 21 to (489.82, 218.25, 164.67) mm, rotated rx 165.67 ry -43.82 rz -104.8 deg; joints [50.471, 29.189, -42.628, -52.248, -64.377, 140.016]
  MoveL 22 to (495.59, 216.52, 164.67) mm, rotated rx 165.67 ry -43.82 rz -104.8 deg; joints [50.245, 28.612, -42.998, -52.284, -64.282, 140.453]
  MoveL 23 to (501.05, 213.4, 164.67) mm, rotated rx 165.67 ry -43.82 rz -104.8 deg; joints [50.138, 27.971, -43.403, -52.389, -64.096, 140.862]
  MoveL 24 to (505.72, 209.03, 164.67) mm, rotated rx 165.67 ry -43.82 rz -104.8 deg; joints [50.174, 27.311, -43.813, -52.564, -63.826, 141.207]
  MoveL 25 to (509.21, 203.76, 164.67) mm, rotated rx 165.67 ry -43.82 rz -104.8 deg; joints [50.355, 26.686, -44.195, -52.802, -63.49, 141.458]
  MoveL 26 to (511.33, 198.05, 164.67) mm, rotated rx 165.67 ry -43.82 rz -104.8 deg; joints [50.662, 26.143, -44.523, -53.081, -63.118, 141.602]
  MoveL 27 to (512.12, 192.37, 164.67) mm, rotated rx 165.67 ry -43.82 rz -104.8 deg; joints [51.058, 25.711, -44.78, -53.378, -62.739, 141.644]
  MoveL 28 to (512.14, 186.87, 164.67) mm, rotated rx 165.67 ry -43.82 rz -104.8 deg; joints [51.495, 25.356, -44.989, -53.679, -62.365, 141.626]
  MoveL 29 to (512.12, 181.36, 164.67) mm, rotated rx 165.67 ry -43.82 rz -104.8 deg; joints [51.939, 25.006, -45.192, -53.982, -61.992, 141.602]
  MoveL 30 to (511.29, 175.68, 164.67) mm, rotated rx 165.67 ry -43.82 rz -104.8 deg; joints [52.455, 24.715, -45.36, -54.308, -61.599, 141.516]
  MoveL 31 to (509.13, 169.97, 164.67) mm, rotated rx 165.67 ry -43.82 rz -104.8 deg; joints [53.061, 24.537, -45.462, -54.65, -61.194, 141.329]
  MoveL 32 to (505.61, 164.72, 164.67) mm, rotated rx 165.67 ry -43.82 rz -104.8 deg; joints [53.717, 24.506, -45.48, -54.979, -60.808, 141.042]
  MoveL 33 to (500.91, 160.38, 164.67) mm, rotated rx 165.67 ry -43.82 rz -104.8 deg; joints [54.367, 24.635, -45.406, -55.261, -60.476, 140.673]
  MoveL 34 to (495.43, 157.3, 164.67) mm, rotated rx 165.67 ry -43.82 rz -104.8 deg; joints [54.953, 24.912, -45.247, -55.47, -60.227, 140.253]
  MoveL 35 to (488.84, 155.47, 164.67) mm, rotated rx 165.67 ry -43.82 rz -104.8 deg; joints [55.493, 25.361, -44.985, -55.605, -60.061, 139.756]
  MoveL 36 to (482.46, 155.19, 164.67) mm, rotated rx 165.67 ry -43.82 rz -104.8 deg; joints [55.883, 25.887, -44.675, -55.642, -60.008, 139.28]
  MoveL 37 to (476.17, 155.19, 164.67) mm, rotated rx 165.67 ry -43.82 rz -104.8 deg; joints [56.237, 26.425, -44.353, -55.655, -59.981, 138.809]
  MoveL 38 to (469.88, 155.19, 164.67) mm, rotated rx 165.67 ry -43.82 rz -104.8 deg; joints [56.585, 26.965, -44.025, -55.659, -59.96, 138.333]
  MoveL 39 to (463.59, 155.19, 164.67) mm, rotated rx 165.67 ry -43.82 rz -104.8 deg; joints [56.927, 27.509, -43.691, -55.656, -59.945, 137.853]
  MoveL 40 to (457.3, 155.19, 164.67) mm, rotated rx 165.67 ry -43.82 rz -104.8 deg; joints [57.262, 28.055, -43.35, -55.644, -59.937, 137.37]
  MoveL 41 to (451.01, 155.19, 164.67) mm, rotated rx 165.67 ry -43.82 rz -104.8 deg; joints [57.591, 28.604, -43.002, -55.625, -59.935, 136.882]
  MoveL 42 to (436.48, 155.19, 164.67) mm, rotated rx 165.67 ry -43.82 rz -104.8 deg; joints [58.33, 29.886, -42.175, -55.552, -59.954, 135.738]
  MoveL 43 to (421.94, 155.19, 164.67) mm, rotated rx 165.67 ry -43.82 rz -104.8 deg; joints [59.039, 31.186, -41.311, -55.44, -60.007, 134.57]
  MoveL 44 to (407.41, 155.4, 164.67) mm, rotated rx 165.67 ry -43.82 rz -104.8 deg; joints [59.703, 32.517, -40.404, -55.28, -60.109, 133.379]
  MoveL 45 to (392.88, 155.08, 164.65) mm, rotated rx 165.67 ry -43.82 rz -104.8 deg; joints [60.383, 33.842, -39.481, -55.111, -60.209, 132.163]
  MoveL 46 to (380.67, 154.12, 163.83) mm, rotated rx 165.67 ry -43.82 rz -104.8 deg; joints [60.986, 34.997, -38.791, -55.015, -60.22, 131.202]
  MoveL 47 to (368.75, 152.58, 161.83) mm, rotated rx 165.67 ry -43.82 rz -104.8 deg; joints [61.604, 36.194, -38.242, -54.983, -60.139, 130.364]
  MoveL 48 to (357.11, 150.48, 158.69) mm, rotated rx 165.67 ry -43.82 rz -104.8 deg; joints [62.235, 37.431, -37.828, -55.012, -59.97, 129.644]
  MoveL 49 to (345.71, 147.84, 154.7) mm, rotated rx 165.67 ry -43.82 rz -104.8 deg; joints [62.879, 38.692, -37.507, -55.083, -59.735, 129.002]
  MoveL 50 to (334.25, 144.58, 151.62) mm, rotated rx 165.67 ry -43.82 rz -104.8 deg; joints [63.556, 39.878, -37.074, -55.105, -59.541, 128.233]
  MoveL 51 to (322.69, 140.7, 149.67) mm, rotated rx 165.67 ry -43.82 rz -104.8 deg; joints [64.264, 40.982, -36.505, -55.062, -59.402, 127.314]
  MoveL 52 to (309.99, 137.13, 148.81) mm, rotated rx 165.67 ry -43.82 rz -104.8 deg; joints [64.971, 42.166, -35.682, -54.886, -59.406, 126.15]
  MoveL 53 to (296.95, 134.79, 148.79) mm, rotated rx 165.67 ry -43.82 rz -104.8 deg; joints [65.581, 43.416, -34.656, -54.575, -59.592, 124.844]
  MoveL 54 to (283.71, 133.72, 148.79) mm, rotated rx 165.67 ry -43.82 rz -104.8 deg; joints [66.088, 44.784, -33.516, -54.176, -59.915, 123.489]
  MoveL 55 to (270.42, 133.93, 148.79) mm, rotated rx 165.67 ry -43.82 rz -104.8 deg; joints [66.489, 46.259, -32.271, -53.702, -60.375, 122.099]
  MoveL 56 to (257.27, 135.41, 148.86) mm, rotated rx 165.67 ry -43.82 rz -104.8 deg; joints [66.784, 47.822, -30.922, -53.164, -60.977, 120.685]
  MoveL 57 to (249.2, 136.96, 149.21) mm, rotated rx 165.67 ry -43.82 rz -104.8 deg; joints [66.916, 48.821, -30.005, -52.791, -61.439, 119.772]
  MoveL 58 to (241.27, 138.98, 149.84) mm, rotated rx 165.67 ry -43.82 rz -104.8 deg; joints [67.008, 49.836, -29.026, -52.391, -61.969, 118.833]
  MoveL 59 to (233.46, 141.48, 150.75) mm, rotated rx 165.67 ry -43.82 rz -104.8 deg; joints [67.064, 50.871, -27.982, -51.969, -62.571, 117.868]
  MoveL 60 to (226.08, 144.9, 151.87) mm, rotated rx 165.67 ry -43.82 rz -104.8 deg; joints [67.044, 51.92, -26.889, -51.526, -63.262, 116.916]
  MoveL 61 to (219.51, 149.71, 153.08) mm, rotated rx 165.67 ry -43.82 rz -104.8 deg; joints [66.909, 52.971, -25.777, -51.074, -64.052, 116.032]
  MoveL 62 to (214.05, 155.71, 154.25) mm, rotated rx 165.67 ry -43.82 rz -104.8 deg; joints [66.668, 53.981, -24.702, -50.639, -64.899, 115.261]
  MoveL 63 to (209.85, 162.72, 155.25) mm, rotated rx 165.67 ry -43.82 rz -104.8 deg; joints [66.329, 54.925, -23.708, -50.238, -65.77, 114.633]
  MoveL 64 to (207.13, 170.42, 155.95) mm, rotated rx 165.67 ry -43.82 rz -104.8 deg; joints [65.91, 55.753, -22.858, -49.894, -66.611, 114.191]
  MoveL 65 to (206.18, 175.85, 156.2) mm, rotated rx 165.67 ry -43.82 rz -104.8 deg; joints [65.59, 56.228, -22.391, -49.7, -67.138, 114.011]
  MoveL 66 to (205.96, 181.36, 156.26) mm, rotated rx 165.67 ry -43.82 rz -104.8 deg; joints [65.245, 56.624, -22.021, -49.539, -67.621, 113.93]
  MoveL 67 to (206.05, 186.88, 156.23) mm, rotated rx 165.67 ry -43.82 rz -104.8 deg; joints [64.893, 56.988, -21.692, -49.392, -68.083, 113.889]
  MoveL 68 to (207.07, 192.25, 155.96) mm, rotated rx 165.67 ry -43.82 rz -104.8 deg; joints [64.525, 57.225, -21.514, -49.292, -68.459, 113.983]
  MoveL 69 to (210.12, 198.87, 155.19) mm, rotated rx 165.67 ry -43.82 rz -104.8 deg; joints [64.018, 57.284, -21.57, -49.243, -68.78, 114.36]
  MoveL 70 to (214.69, 204.51, 154.11) mm, rotated rx 165.67 ry -43.82 rz -104.8 deg; joints [63.525, 57.076, -21.914, -49.276, -68.903, 114.959]
  MoveL 71 to (219.75, 209.66, 153.04) mm, rotated rx 165.67 ry -43.82 rz -104.8 deg; joints [63.045, 56.774, -22.344, -49.333, -68.959, 115.62]
  MoveL 72 to (228.03, 216.62, 151.55) mm, rotated rx 165.67 ry -43.82 rz -104.8 deg; joints [62.345, 56.191, -23.089, -49.442, -68.964, 116.676]
  MoveL 73 to (237.13, 222.66, 150.29) mm, rotated rx 165.67 ry -43.82 rz -104.8 deg; joints [61.669, 55.453, -23.944, -49.578, -68.881, 117.804]
  MoveL 74 to (246.87, 227.62, 149.36) mm, rotated rx 165.67 ry -43.82 rz -104.8 deg; joints [61.028, 54.575, -24.875, -49.735, -68.722, 118.97]
  MoveL 75 to (257.11, 231.44, 148.86) mm, rotated rx 165.67 ry -43.82 rz -104.8 deg; joints [60.432, 53.569, -25.855, -49.909, -68.502, 120.148]
  Establecer velocidad (1000.0 mm/s)
  MoveL 76 to (257.11, 231.44, 148.86) mm, rotated rx 165.67 ry -43.82 rz -104.8 deg; joints [60.432, 53.569, -25.855, -49.909, -68.502, 120.148]
  MoveL 77 to (276.72, 231.44, 246.92) mm, rotated rx 165.67 ry -43.82 rz -104.8 deg; joints [59.721, 46.578, -17.757, -47.738, -74.336, 114.178]
  Establecer velocidad (1000.0 mm/s)
  MoveL 78 to (470.93, 218.86, 311.63) mm, rotated rx 165.67 ry -43.82 rz -104.8 deg; joints [51.551, 21.815, -23.602, -47.354, -76.043, 123.971]
  MoveL 79 to (451.32, 218.86, 213.57) mm, rotated rx 165.67 ry -43.82 rz -104.8 deg; joints [52.664, 28.934, -34.765, -50.432, -67.957, 132.135]
  MoveL 80 to (451.32, 218.86, 213.57) mm, rotated rx 165.67 ry -43.82 rz -104.8 deg; joints [52.664, 28.934, -34.765, -50.432, -67.957, 132.135]
  Establecer velocidad (50.0 mm/s)
  MoveL 81 to (471.17, 217.91, 213.57) mm, rotated rx 165.67 ry -43.82 rz -104.8 deg; joints [51.607, 27.109, -35.804, -50.368, -67.959, 133.592]
  MoveL 82 to (490.86, 215.17, 213.57) mm, rotated rx 165.67 ry -43.82 rz -104.8 deg; joints [50.636, 25.208, -36.831, -50.316, -67.906, 134.983]
  MoveL 83 to (497.27, 213.44, 213.57) mm, rotated rx 165.67 ry -43.82 rz -104.8 deg; joints [50.371, 24.536, -37.179, -50.321, -67.847, 135.419]
  MoveL 84 to (503.1, 210.35, 213.57) mm, rotated rx 165.67 ry -43.82 rz -104.8 deg; joints [50.239, 23.82, -37.543, -50.382, -67.695, 135.794]
  MoveL 85 to (508.17, 206.07, 213.57) mm, rotated rx 165.67 ry -43.82 rz -104.8 deg; joints [50.243, 23.085, -37.907, -50.5, -67.461, 136.095]
  MoveL 86 to (512.17, 200.79, 213.57) mm, rotated rx 165.67 ry -43.82 rz -104.8 deg; joints [50.395, 22.371, -38.251, -50.673, -67.151, 136.301]
  MoveL 87 to (514.69, 194.68, 213.57) mm, rotated rx 165.67 ry -43.82 rz -104.8 deg; joints [50.71, 21.726, -38.555, -50.902, -66.767, 136.387]
  MoveL 88 to (515.43, 188.11, 213.57) mm, rotated rx 165.67 ry -43.82 rz -104.8 deg; joints [51.184, 21.204, -38.795, -51.179, -66.328, 136.337]
  MoveL 89 to (515.11, 181.53, 213.57) mm, rotated rx 165.67 ry -43.82 rz -104.8 deg; joints [51.735, 20.778, -38.987, -51.472, -65.873, 136.209]
  MoveL 90 to (513.23, 175.26, 213.57) mm, rotated rx 165.67 ry -43.82 rz -104.8 deg; joints [52.367, 20.516, -39.104, -51.774, -65.416, 135.975]
  MoveL 91 to (509.75, 169.66, 213.57) mm, rotated rx 165.67 ry -43.82 rz -104.8 deg; joints [53.047, 20.446, -39.135, -52.064, -64.982, 135.643]
  MoveL 92 to (505.15, 164.97, 213.57) mm, rotated rx 165.67 ry -43.82 rz -104.8 deg; joints [53.723, 20.546, -39.091, -52.322, -64.594, 135.248]
  MoveL 93 to (499.81, 161.45, 213.57) mm, rotated rx 165.67 ry -43.82 rz -104.8 deg; joints [54.343, 20.795, -38.979, -52.53, -64.281, 134.825]
  MoveL 94 to (493.83, 159.19, 213.57) mm, rotated rx 165.67 ry -43.82 rz -104.8 deg; joints [54.889, 21.19, -38.801, -52.68, -64.051, 134.381]
  MoveL 95 to (487.59, 158.05, 213.57) mm, rotated rx 165.67 ry -43.82 rz -104.8 deg; joints [55.349, 21.685, -38.574, -52.773, -63.903, 133.938]
  MoveL 96 to (481.3, 157.14, 213.57) mm, rotated rx 165.67 ry -43.82 rz -104.8 deg; joints [55.786, 22.202, -38.331, -52.848, -63.777, 133.492]
  MoveL 97 to (465.19, 155.6, 213.57) mm, rotated rx 165.67 ry -43.82 rz -104.8 deg; joints [56.806, 23.592, -37.656, -52.969, -63.543, 132.351]
  MoveL 98 to (449.01, 155.17, 213.57) mm, rotated rx 165.67 ry -43.82 rz -104.8 deg; joints [57.696, 25.075, -36.9, -52.994, -63.433, 131.199]
  MoveL 99 to (434.31, 155.61, 213.57) mm, rotated rx 165.67 ry -43.82 rz -104.8 deg; joints [58.404, 26.491, -36.144, -52.942, -63.434, 130.141]
  MoveL 100 to (419.75, 157.22, 213.57) mm, rotated rx 165.67 ry -43.82 rz -104.8 deg; joints [58.982, 27.976, -35.316, -52.81, -63.56, 129.087]
  MoveL 101 to (405.48, 159.92, 213.57) mm, rotated rx 165.67 ry -43.82 rz -104.8 deg; joints [59.438, 29.514, -34.424, -52.607, -63.802, 128.042]
  MoveL 102 to (390.94, 159.77, 213.57) mm, rotated rx 165.67 ry -43.82 rz -104.8 deg; joints [60.106, 30.933, -33.569, -52.482, -63.883, 126.912]
  MoveL 103 to (376.41, 159.69, 213.57) mm, rotated rx 165.67 ry -43.82 rz -104.8 deg; joints [60.742, 32.379, -32.669, -52.322, -64.01, 125.755]
  MoveL 104 to (372.08, 159.79, 213.57) mm, rotated rx 165.67 ry -43.82 rz -104.8 deg; joints [60.917, 32.822, -32.388, -52.264, -64.065, 125.407]
  MoveL 105 to (367.77, 160, 213.57) mm, rotated rx 165.67 ry -43.82 rz -104.8 deg; joints [61.082, 33.272, -32.099, -52.199, -64.132, 125.059]
  MoveL 106 to (363.46, 160.37, 213.57) mm, rotated rx 165.67 ry -43.82 rz -104.8 deg; joints [61.232, 33.733, -31.8, -52.127, -64.214, 124.71]
  MoveL 107 to (359.2, 161.07, 213.57) mm, rotated rx 165.67 ry -43.82 rz -104.8 deg; joints [61.354, 34.209, -31.489, -52.042, -64.324, 124.366]
  MoveL 108 to (355.43, 163.13, 213.57) mm, rotated rx 165.67 ry -43.82 rz -104.8 deg; joints [61.355, 34.714, -31.155, -51.916, -64.529, 124.075]
  MoveL 109 to (352.97, 165.76, 213.57) mm, rotated rx 165.67 ry -43.82 rz -104.8 deg; joints [61.26, 35.118, -30.886, -51.791, -64.759, 123.896]
  MoveL 110 to (351.36, 168.97, 213.57) mm, rotated rx 165.67 ry -43.82 rz -104.8 deg; joints [61.089, 35.468, -30.651, -51.659, -65.02, 123.793]
  MoveL 111 to (350.9, 172.52, 213.57) mm, rotated rx 165.67 ry -43.82 rz -104.8 deg; joints [60.847, 35.722, -30.48, -51.534, -65.289, 123.788]
  MoveL 112 to (351.66, 176.05, 213.57) mm, rotated rx 165.67 ry -43.82 rz -104.8 deg; joints [60.561, 35.849, -30.394, -51.429, -65.536, 123.883]
  MoveL 113 to (352.81, 179.48, 213.57) mm, rotated rx 165.67 ry -43.82 rz -104.8 deg; joints [60.264, 35.932, -30.338, -51.331, -65.771, 124.01]
  MoveL 114 to (353.98, 182.91, 213.57) mm, rotated rx 165.67 ry -43.82 rz -104.8 deg; joints [59.968, 36.014, -30.282, -51.234, -66.005, 124.137]
  MoveL 115 to (354.31, 185.66, 213.57) mm, rotated rx 165.67 ry -43.82 rz -104.8 deg; joints [59.757, 36.145, -30.193, -51.147, -66.203, 124.186]
  MoveL 116 to (353.49, 188.44, 213.57) mm, rotated rx 165.67 ry -43.82 rz -104.8 deg; joints [59.593, 36.398, -30.019, -51.045, -66.423, 124.136]
  MoveL 117 to (352.68, 191.22, 213.57) mm, rotated rx 165.67 ry -43.82 rz -104.8 deg; joints [59.428, 36.652, -29.846, -50.943, -66.643, 124.087]
  MoveL 118 to (351.89, 194.01, 213.57) mm, rotated rx 165.67 ry -43.82 rz -104.8 deg; joints [59.264, 36.905, -29.671, -50.842, -66.864, 124.038]
  MoveL 119 to (351.16, 196.81, 213.57) mm, rotated rx 165.67 ry -43.82 rz -104.8 deg; joints [59.097, 37.155, -29.498, -50.742, -67.086, 123.992]
  MoveL 120 to (351.11, 201.63, 213.57) mm, rotated rx 165.67 ry -43.82 rz -104.8 deg; joints [58.761, 37.462, -29.284, -50.585, -67.447, 124.013]
  MoveL 121 to (352.72, 206.18, 213.57) mm, rotated rx 165.67 ry -43.82 rz -104.8 deg; joints [58.375, 37.582, -29.2, -50.458, -67.761, 124.175]
  MoveL 122 to (355.57, 210.09, 213.57) mm, rotated rx 165.67 ry -43.82 rz -104.8 deg; joints [57.982, 37.538, -29.231, -50.365, -68.006, 124.437]
  MoveL 123 to (358.82, 212.66, 213.57) mm, rotated rx 165.67 ry -43.82 rz -104.8 deg; joints [57.662, 37.371, -29.348, -50.316, -68.146, 124.725]
  MoveL 124 to (362.79, 213.91, 213.57) mm, rotated rx 165.67 ry -43.82 rz -104.8 deg; joints [57.402, 37.046, -29.573, -50.316, -68.176, 125.068]
  MoveL 125 to (366.95, 214.46, 213.57) mm, rotated rx 165.67 ry -43.82 rz -104.8 deg; joints [57.178, 36.66, -29.84, -50.337, -68.155, 125.423]
  MoveL 126 to (371.13, 214.8, 213.57) mm, rotated rx 165.67 ry -43.82 rz -104.8 deg; joints [56.967, 36.26, -30.115, -50.363, -68.121, 125.777]
  MoveL 127 to (375.32, 214.97, 213.57) mm, rotated rx 165.67 ry -43.82 rz -104.8 deg; joints [56.765, 35.851, -30.393, -50.392, -68.079, 126.127]
  MoveL 128 to (379.51, 215.02, 213.57) mm, rotated rx 165.67 ry -43.82 rz -104.8 deg; joints [56.569, 35.438, -30.672, -50.422, -68.031, 126.475]
  MoveL 129 to (383.7, 214.99, 213.57) mm, rotated rx 165.67 ry -43.82 rz -104.8 deg; joints [56.377, 35.022, -30.951, -50.453, -67.98, 126.82]
  MoveL 130 to (392.3, 214.76, 213.57) mm, rotated rx 165.67 ry -43.82 rz -104.8 deg; joints [55.988, 34.166, -31.517, -50.515, -67.876, 127.521]
  MoveL 131 to (400.9, 214.49, 213.57) mm, rotated rx 165.67 ry -43.82 rz -104.8 deg; joints [55.594, 33.317, -32.07, -50.568, -67.783, 128.211]
  MoveL 132 to (409.45, 214.97, 213.57) mm, rotated rx 165.67 ry -43.82 rz -104.8 deg; joints [55.139, 32.533, -32.572, -50.583, -67.762, 128.893]
  MoveL 133 to (418.05, 217, 213.57) mm, rotated rx 165.67 ry -43.82 rz -104.8 deg; joints [54.563, 31.857, -32.998, -50.531, -67.865, 129.581]
  MoveL 134 to (423.26, 218.09, 213.57) mm, rotated rx 165.67 ry -43.82 rz -104.8 deg; joints [54.218, 31.444, -33.255, -50.497, -67.925, 129.994]
  MoveL 135 to (427.39, 218.61, 213.57) mm, rotated rx 165.67 ry -43.82 rz -104.8 deg; joints [53.967, 31.096, -33.47, -50.48, -67.95, 130.316]
  MoveL 136 to (430.57, 218.81, 213.57) mm, rotated rx 165.67 ry -43.82 rz -104.8 deg; joints [53.786, 30.816, -33.641, -50.473, -67.957, 130.563]
  MoveL 137 to (433.31, 218.86, 213.57) mm, rotated rx 165.67 ry -43.82 rz -104.8 deg; joints [53.638, 30.568, -33.793, -50.47, -67.955, 130.773]
  MoveL 138 to (436.17, 218.86, 213.57) mm, rotated rx 165.67 ry -43.82 rz -104.8 deg; joints [53.486, 30.306, -33.951, -50.467, -67.952, 130.992]
  MoveL 139 to (438.94, 218.86, 213.57) mm, rotated rx 165.67 ry -43.82 rz -104.8 deg; joints [53.338, 30.052, -34.103, -50.463, -67.949, 131.203]
  MoveL 140 to (442.52, 218.86, 213.57) mm, rotated rx 165.67 ry -43.82 rz -104.8 deg; joints [53.145, 29.727, -34.298, -50.457, -67.949, 131.474]
  MoveL 141 to (446.81, 218.86, 213.57) mm, rotated rx 165.67 ry -43.82 rz -104.8 deg; joints [52.912, 29.34, -34.527, -50.446, -67.951, 131.797]
  MoveL 142 to (451.32, 218.86, 213.57) mm, rotated rx 165.67 ry -43.82 rz -104.8 deg; joints [52.664, 28.934, -34.765, -50.432, -67.957, 132.135]
  Establecer velocidad (1000.0 mm/s)
  MoveL 143 to (451.32, 218.86, 213.57) mm, rotated rx 165.67 ry -43.82 rz -104.8 deg; joints [52.664, 28.934, -34.765, -50.432, -67.957, 132.135]
  MoveL 144 to (470.93, 218.86, 311.63) mm, rotated rx 165.67 ry -43.82 rz -104.8 deg; joints [51.551, 21.815, -23.602, -47.354, -76.043, 123.971]

--- program cerarribder (robot Fanuc LR Mate 200iD/7L) ---
  Suave(1)
  Establecer velocidad (1000.0 mm/s)
  Est. Ref.: RobotiQ 2F-140 Gripper (Mechanism) Base
  Est. herr: Tool 1
  Mostrar Tool 1
  MoveJ 1 to (303.16, 256.16, 250.3) mm, rotated rx -168.7 ry 0.37 rz 88.17 deg; joints [69.758, 40.069, -11.528, -4.201, -67.9, -70.413]
  MoveL 2 to (303.16, 256.16, 250.3) mm, rotated rx -168.7 ry 0.37 rz 88.17 deg; joints [69.758, 40.069, -11.528, -4.201, -67.9, -70.413]
  MoveL 3 to (283.55, 256.16, 152.24) mm, rotated rx -168.7 ry 0.37 rz 88.17 deg; joints [70.263, 45.809, -20.978, -4.46, -58.44, -70.156]
  MoveL 4 to (283.55, 256.16, 152.24) mm, rotated rx -168.7 ry 0.37 rz 88.17 deg; joints [70.263, 45.809, -20.978, -4.46, -58.44, -70.156]
  Establecer velocidad (50.0 mm/s)
  MoveL 5 to (281.45, 256.16, 152.04) mm, rotated rx -168.7 ry 0.37 rz 88.17 deg; joints [70.316, 46.102, -20.777, -4.439, -58.636, -70.232]
  MoveL 6 to (279.36, 256.16, 151.85) mm, rotated rx -168.7 ry 0.37 rz 88.17 deg; joints [70.368, 46.396, -20.573, -4.418, -58.836, -70.307]
  MoveL 7 to (274.03, 256.16, 151.31) mm, rotated rx -168.7 ry 0.37 rz 88.17 deg; joints [70.499, 47.155, -20.05, -4.366, -59.348, -70.498]
  MoveL 8 to (261.94, 256.16, 149.86) mm, rotated rx -168.7 ry 0.37 rz 88.17 deg; joints [70.792, 48.934, -18.827, -4.251, -60.546, -70.921]
  MoveL 9 to (234.64, 256.16, 145.36) mm, rotated rx -168.7 ry 0.37 rz 88.17 deg; joints [71.422, 53.296, -15.823, -4.005, -63.5, -71.846]
  MoveL 10 to (223.99, 256.16, 143.14) mm, rotated rx -168.7 ry 0.37 rz 88.17 deg; joints [71.657, 55.16, -14.523, -3.914, -64.781, -72.197]
  MoveL 11 to (218.06, 256.16, 141.79) mm, rotated rx -168.7 ry 0.37 rz 88.17 deg; joints [71.785, 56.251, -13.756, -3.863, -65.538, -72.391]
  MoveL 12 to (214.74, 256.16, 141) mm, rotated rx -168.7 ry 0.37 rz 88.17 deg; joints [71.857, 56.878, -13.312, -3.835, -65.976, -72.499]
  MoveL 13 to (212.63, 256.16, 140.49) mm, rotated rx -168.7 ry 0.37 rz 88.17 deg; joints [71.901, 57.284, -13.023, -3.818, -66.261, -72.568]
  MoveL 14 to (210.55, 256.16, 139.9) mm, rotated rx -168.7 ry 0.37 rz 88.17 deg; joints [71.945, 57.691, -12.742, -3.801, -66.539, -72.635]
  MoveL 15 to (208.38, 256.16, 137.83) mm, rotated rx -168.7 ry 0.37 rz 88.17 deg; joints [71.991, 58.164, -12.603, -3.788, -66.675, -72.694]
  MoveL 16 to (207.92, 256.16, 136.38) mm, rotated rx -168.7 ry 0.37 rz 88.17 deg; joints [72.001, 58.293, -12.687, -3.788, -66.59, -72.698]
  MoveL 17 to (207.88, 256.16, 134.86) mm, rotated rx -168.7 ry 0.37 rz 88.17 deg; joints [72.002, 58.344, -12.849, -3.793, -66.429, -72.687]
  MoveL 18 to (207.88, 256.16, 128.78) mm, rotated rx -168.7 ry 0.37 rz 88.17 deg; joints [72.002, 58.524, -13.523, -3.812, -65.756, -72.639]
  MoveL 19 to (207.88, 256.16, 116.61) mm, rotated rx -168.7 ry 0.37 rz 88.17 deg; joints [72.002, 58.922, -14.84, -3.853, -64.442, -72.542]
  Establecer velocidad (1000.0 mm/s)
  MoveL 20 to (207.88, 256.16, 116.61) mm, rotated rx -168.7 ry 0.37 rz 88.17 deg; joints [72.002, 58.922, -14.84, -3.853, -64.442, -72.542]
  MoveL 21 to (227.49, 256.16, 214.67) mm, rotated rx -168.7 ry 0.37 rz 88.17 deg; joints [71.58, 53.11, -6.487, -3.721, -72.804, -72.689]
  Establecer velocidad (1000.0 mm/s)
  MoveL 22 to (303.16, 256.16, 250.3) mm, rotated rx -168.7 ry 0.37 rz 88.17 deg; joints [69.758, 40.069, -11.528, -4.201, -67.9, -70.413]
  MoveL 23 to (283.55, 256.16, 152.24) mm, rotated rx -168.7 ry 0.37 rz 88.17 deg; joints [70.263, 45.809, -20.978, -4.46, -58.44, -70.156]
  MoveL 24 to (283.55, 256.16, 152.24) mm, rotated rx -168.7 ry 0.37 rz 88.17 deg; joints [70.263, 45.809, -20.978, -4.46, -58.44, -70.156]
  Establecer velocidad (50.0 mm/s)
  MoveL 25 to (299.11, 256.16, 154.25) mm, rotated rx -168.7 ry 0.37 rz 88.17 deg; joints [69.865, 43.661, -22.342, -4.613, -57.11, -69.593]
  MoveL 26 to (314.45, 256.16, 157.54) mm, rotated rx -168.7 ry 0.37 rz 88.17 deg; joints [69.457, 41.559, -23.435, -4.761, -56.051, -69.037]
  MoveL 27 to (329.49, 256.16, 162.09) mm, rotated rx -168.7 ry 0.37 rz 88.17 deg; joints [69.041, 39.492, -24.264, -4.899, -55.257, -68.494]
  MoveL 28 to (344.09, 256.16, 167.88) mm, rotated rx -168.7 ry 0.37 rz 88.17 deg; joints [68.622, 37.461, -24.83, -5.025, -54.726, -67.97]
  MoveL 29 to (361.89, 256.16, 176.95) mm, rotated rx -168.7 ry 0.37 rz 88.17 deg; joints [68.088, 34.932, -25.176, -5.164, -54.424, -67.341]
  MoveL 30 to (378.65, 256.16, 187.86) mm, rotated rx -168.7 ry 0.37 rz 88.17 deg; joints [67.563, 32.477, -25.111, -5.275, -54.532, -66.766]
  MoveL 31 to (394.18, 256.16, 200.46) mm, rotated rx -168.7 ry 0.37 rz 88.17 deg; joints [67.054, 30.116, -24.65, -5.355, -55.034, -66.256]
  MoveL 32 to (408.29, 256.16, 214.61) mm, rotated rx -168.7 ry 0.37 rz 88.17 deg; joints [66.572, 27.878, -23.811, -5.404, -55.91, -65.821]
  Establecer velocidad (1000.0 mm/s)
  MoveL 33 to (408.29, 256.16, 214.61) mm, rotated rx -168.7 ry 0.37 rz 88.17 deg; joints [66.572, 27.878, -23.811, -5.404, -55.91, -65.821]
  MoveL 34 to (427.9, 256.16, 312.67) mm, rotated rx -168.7 ry 0.37 rz 88.17 deg; joints [65.87, 22.53, -12.532, -4.991, -67.203, -66.225]

--- program talonder (robot Fanuc LR Mate 200iD/7L) ---
  Suave(1)
  Establecer velocidad (1000.0 mm/s)
  Est. Ref.: RobotiQ 2F-140 Gripper (Mechanism) Base
  Est. herr: Tool 1
  Mostrar Tool 1
  MoveJ 1 to (531.86, 166.7, 315.69) mm, rotated rx 173.2 ry -55.45 rz -154.74 deg; joints [53.279, -3.486, -33.006, -72.826, -44.223, 108.835]
  MoveL 2 to (531.86, 166.7, 315.69) mm, rotated rx 173.2 ry -55.45 rz -154.74 deg; joints [53.279, -3.486, -33.006, -72.826, -44.223, 108.835]
  MoveL 3 to (512.24, 166.7, 217.63) mm, rotated rx 173.2 ry -55.45 rz -154.74 deg; joints [54.917, 7.678, -49.066, -91.281, -40.714, 132.222]
  MoveL 4 to (512.24, 166.7, 217.63) mm, rotated rx 173.2 ry -55.45 rz -154.74 deg; joints [54.917, 7.678, -49.066, -91.281, -40.714, 132.222]
  Establecer velocidad (50.0 mm/s)
  MoveL 5 to (514.52, 166.7, 204.48) mm, rotated rx 173.2 ry -55.45 rz -154.74 deg; joints [54.733, 8.994, -51.33, -93.753, -40.931, 135.674]
  MoveL 6 to (517.09, 166.7, 191.38) mm, rotated rx 173.2 ry -55.45 rz -154.74 deg; joints [54.525, 10.364, -53.619, -96.191, -41.256, 139.128]
  MoveL 7 to (519.76, 166.7, 178.31) mm, rotated rx 173.2 ry -55.45 rz -154.74 deg; joints [54.305, 11.807, -55.935, -98.592, -41.68, 142.572]
  MoveL 8 to (521.15, 166.7, 165.64) mm, rotated rx 173.2 ry -55.45 rz -154.74 deg; joints [54.189, 13.385, -58.162, -100.93, -42.119, 145.842]
  MoveL 9 to (521.11, 166.7, 152.93) mm, rotated rx 173.2 ry -55.45 rz -154.74 deg; joints [54.193, 15.154, -60.355, -103.286, -42.578, 149.026]
  MoveL 10 to (519.65, 166.7, 140.38) mm, rotated rx 173.2 ry -55.45 rz -154.74 deg; joints [54.314, 17.06, -62.452, -105.6, -43.045, 152.035]
  MoveL 11 to (516.78, 166.7, 128.05) mm, rotated rx 173.2 ry -55.45 rz -154.74 deg; joints [54.55, 19.076, -64.422, -107.848, -43.511, 154.833]
  Establecer velocidad (1000.0 mm/s)
  MoveL 12 to (516.78, 166.7, 128.05) mm, rotated rx 173.2 ry -55.45 rz -154.74 deg; joints [54.55, 19.076, -64.422, -107.848, -43.511, 154.833]
  MoveL 13 to (536.39, 166.7, 226.11) mm, rotated rx 173.2 ry -55.45 rz -154.74 deg; joints [52.882, 4.393, -47.97, -88.516, -42.064, 130.569]

--- program iman izquierdo (robot Fanuc LR Mate 200iD/7L) ---
  Est. Ref.: iman izquierdo
  Est. herr: Tool 1
  MoveJ (Target 1)
  MoveL (Target 2)
  MoveL (Target 3)
  Llamar close
  Adjuntar a Tool 1
  MoveL (Target 4)
  MoveJ (Target 5)
  MoveL (Target 6)
  Llamar open
  Separar de Tool 1
  MoveJ (Target 5)

--- program iman derecho (robot Fanuc LR Mate 200iD/7L) ---
  Est. Ref.: iman derecho
  Est. herr: Tool 1
  MoveJ (Target 1)
  MoveL (Target 2)
  MoveL (Target 3)
  Llamar close
  Adjuntar a Tool 1
  MoveL (Target 4)
  MoveJ (Target 5)
  MoveL (Target 6)
  Llamar open
  Separar de Tool 1
  MoveJ (Target 5)

--- program dejar iman izquierdo (robot Fanuc LR Mate 200iD/7L) ---
  Est. Ref.: iman izquierdo
  Est. herr: Tool 1
  MoveJ (Target 6)
  Llamar close
  Adjuntar a Tool 1
  MoveL (Target 5)
  MoveL (Target 4)
  MoveL (Target 3)
  MoveL (Target 2)
  Llamar open
  Separar de Tool 1
  MoveL (Target 1)

--- program dejar iman derecho (robot Fanuc LR Mate 200iD/7L) ---
  Est. Ref.: iman derecho
  Est. herr: Tool 1
  MoveJ (Target 6)
  Llamar open
  Adjuntar a Tool 1
  MoveL (Target 5)
  MoveL (Target 4)
  MoveL (Target 3)
  MoveL (Target 2)
  Llamar open
  Separar de Tool 1
  MoveL (Target 1)

--- program platizch (robot Fanuc LR Mate 200iD/7L) ---
  Suave(1)
  Establecer velocidad (1000.0 mm/s)
  Est. Ref.: RobotiQ 2F-140 Gripper (Mechanism) Base
  Est. herr: Tool 1
  Mostrar Tool 1
  MoveJ 1 to (276.49, 139.55, 274.86) mm, rotated rx 150.39 ry -54.39 rz -78.94 deg; joints [57.109, 41.788, -24.817, -58.793, -84.834, 135.304]
  MoveL 2 to (276.49, 139.55, 274.86) mm, rotated rx 150.39 ry -54.39 rz -78.94 deg; joints [57.109, 41.788, -24.817, -58.793, -84.834, 135.304]
  MoveL 3 to (256.88, 139.55, 176.81) mm, rotated rx 150.39 ry -54.39 rz -78.94 deg; joints [57.917, 49.529, -33.108, -60.089, -80.004, 142.141]
  MoveL 4 to (256.88, 139.55, 176.81) mm, rotated rx 150.39 ry -54.39 rz -78.94 deg; joints [57.917, 49.529, -33.108, -60.089, -80.004, 142.141]
  Establecer velocidad (50.0 mm/s)
  MoveL 5 to (266.27, 140.34, 176.8) mm, rotated rx 150.39 ry -54.39 rz -78.94 deg; joints [57.484, 48.614, -33.931, -60.009, -79.906, 143.048]
  MoveL 6 to (275.71, 140.33, 176.8) mm, rotated rx 150.39 ry -54.39 rz -78.94 deg; joints [57.091, 47.665, -34.78, -59.948, -79.762, 143.96]
  MoveL 7 to (285.12, 139.52, 176.8) mm, rotated rx 150.39 ry -54.39 rz -78.94 deg; joints [56.745, 46.689, -35.647, -59.911, -79.572, 144.867]
  MoveL 8 to (294.39, 137.92, 176.8) mm, rotated rx 150.39 ry -54.39 rz -78.94 deg; joints [56.448, 45.696, -36.522, -59.899, -79.341, 145.759]
  MoveL 9 to (303.47, 135.55, 177.24) mm, rotated rx 150.39 ry -54.39 rz -78.94 deg; joints [56.204, 44.662, -37.357, -59.909, -79.091, 146.594]
  MoveL 10 to (312.83, 132.4, 178.57) mm, rotated rx 150.39 ry -54.39 rz -78.94 deg; joints [55.994, 43.505, -38.142, -59.929, -78.841, 147.372]
  MoveL 11 to (322.11, 129.63, 180.81) mm, rotated rx 150.39 ry -54.39 rz -78.94 deg; joints [55.756, 42.328, -38.783, -59.91, -78.682, 148.032]
  MoveL 12 to (331.3, 127.37, 183.95) mm, rotated rx 150.39 ry -54.39 rz -78.94 deg; joints [55.48, 41.134, -39.271, -59.842, -78.622, 148.572]
  MoveL 13 to (340.63, 125.56, 186.74) mm, rotated rx 150.39 ry -54.39 rz -78.94 deg; joints [55.16, 39.989, -39.754, -59.748, -78.592, 149.125]
  MoveL 14 to (350.19, 124.18, 188.6) mm, rotated rx 150.39 ry -54.39 rz -78.94 deg; joints [54.789, 38.93, -40.304, -59.634, -78.56, 149.756]
  MoveL 15 to (359.98, 123.28, 189.53) mm, rotated rx 150.39 ry -54.39 rz -78.94 deg; joints [54.363, 37.96, -40.925, -59.499, -78.524, 150.469]
  MoveL 16 to (370.64, 122.86, 189.63) mm, rotated rx 150.39 ry -54.39 rz -78.94 deg; joints [53.848, 37.024, -41.649, -59.326, -78.489, 151.306]
  MoveL 17 to (381.3, 123.03, 189.63) mm, rotated rx 150.39 ry -54.39 rz -78.94 deg; joints [53.276, 36.144, -42.336, -59.107, -78.502, 152.13]
  MoveL 18 to (391.96, 123.03, 189.63) mm, rotated rx 150.39 ry -54.39 rz -78.94 deg; joints [52.701, 35.269, -43.012, -58.88, -78.516, 152.944]
  MoveL 19 to (402.63, 123.03, 189.63) mm, rotated rx 150.39 ry -54.39 rz -78.94 deg; joints [52.11, 34.406, -43.67, -58.634, -78.543, 153.745]
  MoveL 20 to (413.29, 123.03, 189.63) mm, rotated rx 150.39 ry -54.39 rz -78.94 deg; joints [51.503, 33.557, -44.31, -58.369, -78.581, 154.534]
  MoveL 21 to (419.95, 123.03, 189.63) mm, rotated rx 150.39 ry -54.39 rz -78.94 deg; joints [51.116, 33.033, -44.7, -58.193, -78.61, 155.021]
  MoveL 22 to (426.62, 123.03, 189.63) mm, rotated rx 150.39 ry -54.39 rz -78.94 deg; joints [50.722, 32.514, -45.084, -58.01, -78.645, 155.504]
  MoveL 23 to (433.28, 123.03, 189.63) mm, rotated rx 150.39 ry -54.39 rz -78.94 deg; joints [50.321, 31.999, -45.461, -57.819, -78.683, 155.983]
  MoveL 24 to (440.01, 122.83, 189.63) mm, rotated rx 150.39 ry -54.39 rz -78.94 deg; joints [49.923, 31.472, -45.844, -57.63, -78.714, 156.465]
  MoveL 25 to (444.67, 121.68, 189.63) mm, rotated rx 150.39 ry -54.39 rz -78.94 deg; joints [49.719, 31.044, -46.153, -57.55, -78.669, 156.808]
  MoveL 26 to (449.17, 119.42, 189.63) mm, rotated rx 150.39 ry -54.39 rz -78.94 deg; joints [49.604, 30.559, -46.499, -57.534, -78.549, 157.15]
  MoveL 27 to (453.11, 116.1, 189.63) mm, rotated rx 150.39 ry -54.39 rz -78.94 deg; joints [49.6, 30.049, -46.86, -57.594, -78.358, 157.462]
  MoveL 28 to (456.16, 111.98, 189.63) mm, rotated rx 150.39 ry -54.39 rz -78.94 deg; joints [49.715, 29.556, -47.206, -57.73, -78.107, 157.717]
  MoveL 29 to (458.14, 107.42, 189.63) mm, rotated rx 150.39 ry -54.39 rz -78.94 deg; joints [49.936, 29.118, -47.51, -57.931, -77.818, 157.899]
  MoveL 30 to (459.01, 102.8, 189.63) mm, rotated rx 150.39 ry -54.39 rz -78.94 deg; joints [50.234, 28.76, -47.756, -58.174, -77.517, 158.004]
  MoveL 31 to (459.08, 98.35, 189.63) mm, rotated rx 150.39 ry -54.39 rz -78.94 deg; joints [50.576, 28.476, -47.951, -58.437, -77.22, 158.05]
  MoveL 32 to (459.08, 93.9, 189.63) mm, rotated rx 150.39 ry -54.39 rz -78.94 deg; joints [50.925, 28.2, -48.139, -58.705, -76.923, 158.09]
  MoveL 33 to (458.65, 89.36, 189.63) mm, rotated rx 150.39 ry -54.39 rz -78.94 deg; joints [51.312, 27.954, -48.305, -58.996, -76.616, 158.1]
  MoveL 34 to (457.17, 84.73, 189.63) mm, rotated rx 150.39 ry -54.39 rz -78.94 deg; joints [51.777, 27.785, -48.419, -59.329, -76.293, 158.037]
  MoveL 35 to (454.58, 80.37, 189.63) mm, rotated rx 150.39 ry -54.39 rz -78.94 deg; joints [52.292, 27.723, -48.461, -59.681, -75.977, 157.896]
  MoveL 36 to (450.99, 76.66, 189.63) mm, rotated rx 150.39 ry -54.39 rz -78.94 deg; joints [52.817, 27.781, -48.422, -60.02, -75.696, 157.68]
  MoveL 37 to (446.68, 73.92, 189.63) mm, rotated rx 150.39 ry -54.39 rz -78.94 deg; joints [53.305, 27.957, -48.303, -60.317, -75.473, 157.408]
  MoveL 38 to (442.05, 72.28, 189.63) mm, rotated rx 150.39 ry -54.39 rz -78.94 deg; joints [53.719, 28.227, -48.12, -60.549, -75.323, 157.102]
  MoveL 39 to (435.97, 71.72, 189.63) mm, rotated rx 150.39 ry -54.39 rz -78.94 deg; joints [54.127, 28.676, -47.814, -60.747, -75.236, 156.688]
  MoveL 40 to (430.05, 71.72, 189.63) mm, rotated rx 150.39 ry -54.39 rz -78.94 deg; joints [54.473, 29.149, -47.488, -60.898, -75.191, 156.276]
  MoveL 41 to (424.12, 71.72, 189.63) mm, rotated rx 150.39 ry -54.39 rz -78.94 deg; joints [54.814, 29.625, -47.157, -61.042, -75.149, 155.861]
  MoveL 42 to (418.2, 71.72, 189.63) mm, rotated rx 150.39 ry -54.39 rz -78.94 deg; joints [55.149, 30.104, -46.821, -61.179, -75.112, 155.442]
  MoveL 43 to (412.28, 71.72, 189.63) mm, rotated rx 150.39 ry -54.39 rz -78.94 deg; joints [55.479, 30.586, -46.479, -61.31, -75.078, 155.019]
  MoveL 44 to (406.35, 71.72, 189.63) mm, rotated rx 150.39 ry -54.39 rz -78.94 deg; joints [55.803, 31.071, -46.132, -61.435, -75.047, 154.593]
  MoveL 45 to (394.62, 71.72, 189.63) mm, rotated rx 150.39 ry -54.39 rz -78.94 deg; joints [56.429, 32.041, -45.43, -61.663, -74.998, 153.739]
  MoveL 46 to (382.89, 71.72, 189.63) mm, rotated rx 150.39 ry -54.39 rz -78.94 deg; joints [57.035, 33.025, -44.706, -61.866, -74.963, 152.869]
  MoveL 47 to (371.17, 71.32, 189.63) mm, rotated rx 150.39 ry -54.39 rz -78.94 deg; joints [57.652, 34, -43.977, -62.069, -74.916, 151.987]
  MoveL 48 to (359.5, 70.13, 189.51) mm, rotated rx 150.39 ry -54.39 rz -78.94 deg; joints [58.309, 34.951, -43.276, -62.295, -74.823, 151.115]
  MoveL 49 to (349.79, 68.52, 188.55) mm, rotated rx 150.39 ry -54.39 rz -78.94 deg; joints [58.889, 35.792, -42.796, -62.521, -74.669, 150.471]
  MoveL 50 to (340.32, 66.39, 186.66) mm, rotated rx 150.39 ry -54.39 rz -78.94 deg; joints [59.485, 36.667, -42.436, -62.78, -74.445, 149.93]
  MoveL 51 to (331.08, 63.88, 183.87) mm, rotated rx 150.39 ry -54.39 rz -78.94 deg; joints [60.086, 37.582, -42.188, -63.066, -74.163, 149.49]
  MoveL 52 to (321.89, 61.73, 180.75) mm, rotated rx 150.39 ry -54.39 rz -78.94 deg; joints [60.645, 38.547, -41.941, -63.324, -73.903, 149.066]
  MoveL 53 to (312.46, 60.05, 178.5) mm, rotated rx 150.39 ry -54.39 rz -78.94 deg; joints [61.168, 39.496, -41.542, -63.518, -73.733, 148.513]
  MoveL 54 to (302.79, 58.84, 177.18) mm, rotated rx 150.39 ry -54.39 rz -78.94 deg; joints [61.654, 40.428, -40.988, -63.645, -73.653, 147.827]
  MoveL 55 to (293.95, 58.19, 176.8) mm, rotated rx 150.39 ry -54.39 rz -78.94 deg; joints [62.054, 41.25, -40.359, -63.701, -73.66, 147.099]
  MoveL 56 to (285.04, 57.97, 176.8) mm, rotated rx 150.39 ry -54.39 rz -78.94 deg; joints [62.416, 42.082, -39.651, -63.713, -73.725, 146.31]
  MoveL 57 to (276.13, 57.97, 176.8) mm, rotated rx 150.39 ry -54.39 rz -78.94 deg; joints [62.754, 42.939, -38.917, -63.702, -73.815, 145.504]
  MoveL 58 to (267.23, 58.45, 176.8) mm, rotated rx 150.39 ry -54.39 rz -78.94 deg; joints [63.05, 43.833, -38.146, -63.656, -73.949, 144.678]
  MoveL 59 to (258.45, 59.95, 176.8) mm, rotated rx 150.39 ry -54.39 rz -78.94 deg; joints [63.261, 44.782, -37.322, -63.554, -74.166, 143.832]
  MoveL 60 to (249.91, 62.45, 176.97) mm, rotated rx 150.39 ry -54.39 rz -78.94 deg; joints [63.389, 45.762, -36.437, -63.395, -74.47, 142.963]
  MoveL 61 to (241.75, 65.89, 177.51) mm, rotated rx 150.39 ry -54.39 rz -78.94 deg; joints [63.434, 46.744, -35.486, -63.184, -74.865, 142.065]
  MoveL 62 to (234.01, 70.27, 178.37) mm, rotated rx 150.39 ry -54.39 rz -78.94 deg; joints [63.399, 47.729, -34.476, -62.928, -75.348, 141.147]
  MoveL 63 to (226.89, 75.45, 179.47) mm, rotated rx 150.39 ry -54.39 rz -78.94 deg; joints [63.288, 48.701, -33.438, -62.64, -75.904, 140.238]
  MoveL 64 to (222.93, 78.92, 180.21) mm, rotated rx 150.39 ry -54.39 rz -78.94 deg; joints [63.188, 49.275, -32.809, -62.457, -76.269, 139.702]
  MoveL 65 to (219.21, 82.66, 181) mm, rotated rx 150.39 ry -54.39 rz -78.94 deg; joints [63.063, 49.846, -32.177, -62.267, -76.656, 139.177]
  MoveL 66 to (215.77, 86.7, 181.79) mm, rotated rx 150.39 ry -54.39 rz -78.94 deg; joints [62.91, 50.412, -31.546, -62.07, -77.065, 138.665]
  MoveL 67 to (213.2, 91.34, 182.44) mm, rotated rx 150.39 ry -54.39 rz -78.94 deg; joints [62.689, 50.934, -30.977, -61.862, -77.499, 138.242]
  MoveL 68 to (211.86, 96.49, 182.79) mm, rotated rx 150.39 ry -54.39 rz -78.94 deg; joints [62.396, 51.372, -30.527, -61.652, -77.934, 137.959]
  MoveL 69 to (211.69, 102.45, 182.84) mm, rotated rx 150.39 ry -54.39 rz -78.94 deg; joints [62.012, 51.752, -30.176, -61.426, -78.393, 137.804]
  MoveL 70 to (212.15, 108.39, 182.71) mm, rotated rx 150.39 ry -54.39 rz -78.94 deg; joints [61.61, 52.076, -29.901, -61.21, -78.83, 137.729]
  MoveL 71 to (213.66, 114.12, 182.32) mm, rotated rx 150.39 ry -54.39 rz -78.94 deg; joints [61.187, 52.288, -29.767, -61.011, -79.216, 137.789]
  MoveL 72 to (216.15, 119.45, 181.7) mm, rotated rx 150.39 ry -54.39 rz -78.94 deg; joints [60.756, 52.381, -29.774, -60.832, -79.539, 137.981]
  MoveL 73 to (219.54, 124.26, 180.92) mm, rotated rx 150.39 ry -54.39 rz -78.94 deg; joints [60.326, 52.351, -29.919, -60.675, -79.794, 138.294]
  MoveL 74 to (223.71, 128.37, 180.06) mm, rotated rx 150.39 ry -54.39 rz -78.94 deg; joints [59.911, 52.198, -30.189, -60.54, -79.975, 138.712]
  MoveL 75 to (228.54, 131.69, 179.19) mm, rotated rx 150.39 ry -54.39 rz -78.94 deg; joints [59.52, 51.924, -30.57, -60.43, -80.08, 139.218]
  MoveL 76 to (233.89, 134.1, 178.39) mm, rotated rx 150.39 ry -54.39 rz -78.94 deg; joints [59.165, 51.537, -31.044, -60.346, -80.111, 139.79]
  MoveL 77 to (239.52, 135.92, 177.72) mm, rotated rx 150.39 ry -54.39 rz -78.94 deg; joints [58.834, 51.081, -31.56, -60.277, -80.101, 140.387]
  MoveL 78 to (245.22, 137.43, 177.23) mm, rotated rx 150.39 ry -54.39 rz -78.94 deg; joints [58.515, 50.595, -32.077, -60.211, -80.08, 140.979]
  MoveL 79 to (251.01, 138.64, 176.92) mm, rotated rx 150.39 ry -54.39 rz -78.94 deg; joints [58.209, 50.078, -32.593, -60.148, -80.047, 141.564]
  MoveL 80 to (256.88, 139.55, 176.81) mm, rotated rx 150.39 ry -54.39 rz -78.94 deg; joints [57.917, 49.529, -33.108, -60.089, -80.004, 142.141]
  Establecer velocidad (1000.0 mm/s)
  MoveL 81 to (256.88, 139.55, 176.81) mm, rotated rx 150.39 ry -54.39 rz -78.94 deg; joints [57.917, 49.529, -33.108, -60.089, -80.004, 142.141]
  MoveL 82 to (276.49, 139.55, 274.86) mm, rotated rx 150.39 ry -54.39 rz -78.94 deg; joints [57.109, 41.788, -24.817, -58.793, -84.834, 135.304]
  Establecer velocidad (1000.0 mm/s)
  MoveL 83 to (429.55, 71.57, 327.09) mm, rotated rx 150.39 ry -54.39 rz -78.94 deg; joints [54.514, 19.004, -30.081, -58.15, -84.045, 141.022]
  MoveL 84 to (409.94, 71.57, 229.03) mm, rotated rx 150.39 ry -54.39 rz -78.94 deg; joints [55.619, 27.475, -41.595, -60.35, -77.372, 150.578]
  MoveL 85 to (409.94, 71.57, 229.03) mm, rotated rx 150.39 ry -54.39 rz -78.94 deg; joints [55.619, 27.475, -41.595, -60.35, -77.372, 150.578]
  Establecer velocidad (50.0 mm/s)
  MoveL 86 to (426.07, 72.34, 229.03) mm, rotated rx 150.39 ry -54.39 rz -78.94 deg; joints [54.652, 26.126, -42.392, -59.936, -77.598, 151.652]
  MoveL 87 to (442.07, 74.58, 229.03) mm, rotated rx 150.39 ry -54.39 rz -78.94 deg; joints [53.53, 24.901, -43.091, -59.395, -77.956, 152.695]
  MoveL 88 to (447.27, 76.02, 229.03) mm, rotated rx 150.39 ry -54.39 rz -78.94 deg; joints [53.097, 24.553, -43.285, -59.168, -78.128, 153.03]
  MoveL 89 to (451.99, 78.57, 229.03) mm, rotated rx 150.39 ry -54.39 rz -78.94 deg; joints [52.599, 24.32, -43.413, -58.888, -78.373, 153.334]
  MoveL 90 to (456.08, 82.09, 229.03) mm, rotated rx 150.39 ry -54.39 rz -78.94 deg; joints [52.058, 24.206, -43.476, -58.568, -78.676, 153.596]
  MoveL 91 to (459.27, 86.43, 229.03) mm, rotated rx 150.39 ry -54.39 rz -78.94 deg; joints [51.506, 24.224, -43.466, -58.228, -79.022, 153.802]
  MoveL 92 to (461.24, 91.43, 229.03) mm, rotated rx 150.39 ry -54.39 rz -78.94 deg; joints [50.981, 24.392, -43.374, -57.891, -79.395, 153.927]
  MoveL 93 to (461.75, 96.76, 229.03) mm, rotated rx 150.39 ry -54.39 rz -78.94 deg; joints [50.528, 24.704, -43.201, -57.586, -79.766, 153.957]
  MoveL 94 to (461.6, 101.04, 229.03) mm, rotated rx 150.39 ry -54.39 rz -78.94 deg; joints [50.204, 25.003, -43.034, -57.362, -80.055, 153.943]
  MoveL 95 to (460.62, 105.15, 229.03) mm, rotated rx 150.39 ry -54.39 rz -78.94 deg; joints [49.95, 25.359, -42.833, -57.177, -80.321, 153.874]
  MoveL 96 to (458.82, 109, 229.03) mm, rotated rx 150.39 ry -54.39 rz -78.94 deg; joints [49.771, 25.765, -42.601, -57.035, -80.557, 153.749]
  MoveL 97 to (456.31, 112.39, 229.03) mm, rotated rx 150.39 ry -54.39 rz -78.94 deg; joints [49.675, 26.197, -42.351, -56.942, -80.752, 153.576]
  MoveL 98 to (453.24, 115.32, 229.03) mm, rotated rx 150.39 ry -54.39 rz -78.94 deg; joints [49.651, 26.644, -42.09, -56.892, -80.91, 153.364]
  MoveL 99 to (448.52, 118.3, 229.03) mm, rotated rx 150.39 ry -54.39 rz -78.94 deg; joints [49.727, 27.226, -41.744, -56.892, -81.051, 153.039]
  MoveL 100 to (443.2, 120.06, 229.03) mm, rotated rx 150.39 ry -54.39 rz -78.94 deg; joints [49.929, 27.775, -41.414, -56.97, -81.105, 152.676]
  MoveL 101 to (437.68, 120.98, 229.03) mm, rotated rx 150.39 ry -54.39 rz -78.94 deg; joints [50.202, 28.286, -41.102, -57.091, -81.102, 152.298]
  MoveL 102 to (432.14, 121.73, 229.03) mm, rotated rx 150.39 ry -54.39 rz -78.94 deg; joints [50.485, 28.789, -40.791, -57.217, -81.091, 151.916]
  MoveL 103 to (426.57, 122.3, 229.03) mm, rotated rx 150.39 ry -54.39 rz -78.94 deg; joints [50.777, 29.286, -40.481, -57.348, -81.073, 151.531]
  MoveL 104 to (420.99, 122.72, 229.03) mm, rotated rx 150.39 ry -54.39 rz -78.94 deg; joints [51.077, 29.775, -40.171, -57.482, -81.046, 151.142]
  MoveL 105 to (407.8, 123.06, 229.03) mm, rotated rx 150.39 ry -54.39 rz -78.94 deg; joints [51.816, 30.901, -39.446, -57.809, -80.956, 150.214]
  MoveL 106 to (394.62, 122.59, 229.03) mm, rotated rx 150.39 ry -54.39 rz -78.94 deg; joints [52.587, 31.992, -38.726, -58.147, -80.829, 149.275]
  MoveL 107 to (386.84, 121.75, 229.03) mm, rotated rx 150.39 ry -54.39 rz -78.94 deg; joints [53.071, 32.608, -38.313, -58.359, -80.725, 148.717]
  MoveL 108 to (379.18, 120.43, 229.03) mm, rotated rx 150.39 ry -54.39 rz -78.94 deg; joints [53.574, 33.191, -37.917, -58.58, -80.594, 148.165]
  MoveL 109 to (371.55, 119.23, 229.03) mm, rotated rx 150.39 ry -54.39 rz -78.94 deg; joints [54.06, 33.787, -37.508, -58.785, -80.479, 147.609]
  MoveL 110 to (363.79, 119.31, 229.03) mm, rotated rx 150.39 ry -54.39 rz -78.94 deg; joints [54.452, 34.484, -37.024, -58.926, -80.462, 147.025]
  MoveL 111 to (356.03, 119.43, 229.03) mm, rotated rx 150.39 ry -54.39 rz -78.94 deg; joints [54.834, 35.192, -36.526, -59.057, -80.456, 146.432]
  MoveL 112 to (348.27, 119.41, 229.03) mm, rotated rx 150.39 ry -54.39 rz -78.94 deg; joints [55.218, 35.898, -36.023, -59.185, -80.449, 145.833]
  MoveL 113 to (344.75, 119.31, 229.03) mm, rotated rx 150.39 ry -54.39 rz -78.94 deg; joints [55.397, 36.215, -35.796, -59.244, -80.441, 145.56]
  MoveL 114 to (341.23, 119.1, 229.03) mm, rotated rx 150.39 ry -54.39 rz -78.94 deg; joints [55.581, 36.528, -35.57, -59.306, -80.427, 145.286]
  MoveL 115 to (337.72, 118.75, 229.03) mm, rotated rx 150.39 ry -54.39 rz -78.94 deg; joints [55.773, 36.832, -35.349, -59.372, -80.405, 145.012]
  MoveL 116 to (334.29, 117.91, 229.03) mm, rotated rx 150.39 ry -54.39 rz -78.94 deg; joints [55.994, 37.099, -35.155, -59.456, -80.349, 144.749]
  MoveL 117 to (331.42, 115.87, 229.03) mm, rotated rx 150.39 ry -54.39 rz -78.94 deg; joints [56.272, 37.24, -35.052, -59.581, -80.205, 144.542]
  MoveL 118 to (329.65, 113.51, 229.03) mm, rotated rx 150.39 ry -54.39 rz -78.94 deg; joints [56.52, 37.259, -35.038, -59.703, -80.037, 144.426]
  MoveL 119 to (328.69, 110.73, 229.03) mm, rotated rx 150.39 ry -54.39 rz -78.94 deg; joints [56.761, 37.177, -35.098, -59.833, -79.837, 144.378]
  MoveL 120 to (328.75, 107.79, 229.03) mm, rotated rx 150.39 ry -54.39 rz -78.94 deg; joints [56.966, 36.989, -35.235, -59.957, -79.623, 144.413]
  MoveL 121 to (330.08, 103.57, 229.03) mm, rotated rx 150.39 ry -54.39 rz -78.94 deg; joints [57.205, 36.606, -35.514, -60.122, -79.315, 144.559]
  MoveL 122 to (331.52, 99.39, 229.03) mm, rotated rx 150.39 ry -54.39 rz -78.94 deg; joints [57.438, 36.216, -35.795, -60.287, -79.011, 144.712]
  MoveL 123 to (331.08, 97.51, 229.03) mm, rotated rx 150.39 ry -54.39 rz -78.94 deg; joints [57.594, 36.145, -35.846, -60.375, -78.876, 144.694]
  MoveL 124 to (330.52, 95.62, 229.03) mm, rotated rx 150.39 ry -54.39 rz -78.94 deg; joints [57.755, 36.084, -35.89, -60.464, -78.74, 144.666]
  MoveL 125 to (329.98, 93.74, 229.03) mm, rotated rx 150.39 ry -54.39 rz -78.94 deg; joints [57.917, 36.023, -35.933, -60.553, -78.605, 144.639]
  MoveL 126 to (329.45, 91.84, 229.03) mm, rotated rx 150.39 ry -54.39 rz -78.94 deg; joints [58.079, 35.962, -35.977, -60.643, -78.469, 144.613]
  MoveL 127 to (328.92, 89.95, 229.03) mm, rotated rx 150.39 ry -54.39 rz -78.94 deg; joints [58.24, 35.9, -36.022, -60.733, -78.333, 144.587]
  MoveL 128 to (328.62, 88.02, 229.03) mm, rotated rx 150.39 ry -54.39 rz -78.94 deg; joints [58.395, 35.815, -36.082, -60.822, -78.195, 144.579]
  MoveL 129 to (329.08, 84.17, 229.03) mm, rotated rx 150.39 ry -54.39 rz -78.94 deg; joints [58.656, 35.548, -36.273, -60.99, -77.917, 144.644]
  MoveL 130 to (330.77, 80.67, 229.03) mm, rotated rx 150.39 ry -54.39 rz -78.94 deg; joints [58.839, 35.186, -36.53, -61.132, -77.664, 144.802]
  MoveL 131 to (333.33, 77.75, 229.03) mm, rotated rx 150.39 ry -54.39 rz -78.94 deg; joints [58.941, 34.776, -36.819, -61.24, -77.454, 145.02]
  MoveL 132 to (336.71, 75.85, 229.03) mm, rotated rx 150.39 ry -54.39 rz -78.94 deg; joints [58.931, 34.349, -37.118, -61.293, -77.317, 145.293]
  MoveL 133 to (340.54, 75.21, 229.03) mm, rotated rx 150.39 ry -54.39 rz -78.94 deg; joints [58.805, 33.952, -37.394, -61.282, -77.272, 145.59]
  MoveL 134 to (344.42, 74.86, 229.03) mm, rotated rx 150.39 ry -54.39 rz -78.94 deg; joints [58.654, 33.568, -37.658, -61.256, -77.25, 145.887]
  MoveL 135 to (348.31, 74.69, 229.03) mm, rotated rx 150.39 ry -54.39 rz -78.94 deg; joints [58.487, 33.196, -37.913, -61.219, -77.243, 146.181]
  MoveL 136 to (352.21, 74.64, 229.03) mm, rotated rx 150.39 ry -54.39 rz -78.94 deg; joints [58.308, 32.833, -38.161, -61.173, -77.247, 146.473]
  MoveL 137 to (356.1, 74.69, 229.03) mm, rotated rx 150.39 ry -54.39 rz -78.94 deg; joints [58.121, 32.476, -38.402, -61.121, -77.26, 146.762]
  MoveL 138 to (360.46, 74.8, 229.03) mm, rotated rx 150.39 ry -54.39 rz -78.94 deg; joints [57.904, 32.082, -38.666, -61.056, -77.281, 147.084]
  MoveL 139 to (364.82, 74.95, 229.03) mm, rotated rx 150.39 ry -54.39 rz -78.94 deg; joints [57.682, 31.692, -38.925, -60.987, -77.306, 147.402]
  MoveL 140 to (369.18, 75.09, 229.03) mm, rotated rx 150.39 ry -54.39 rz -78.94 deg; joints [57.458, 31.303, -39.182, -60.916, -77.334, 147.719]
  MoveL 141 to (373.54, 75.18, 229.03) mm, rotated rx 150.39 ry -54.39 rz -78.94 deg; joints [57.235, 30.914, -39.437, -60.843, -77.361, 148.033]
  MoveL 142 to (377.83, 74.36, 229.03) mm, rotated rx 150.39 ry -54.39 rz -78.94 deg; joints [57.084, 30.481, -39.718, -60.815, -77.325, 148.343]
  MoveL 143 to (382.15, 73.31, 229.03) mm, rotated rx 150.39 ry -54.39 rz -78.94 deg; joints [56.947, 30.032, -40.006, -60.796, -77.276, 148.653]
  MoveL 144 to (386.89, 72.24, 229.03) mm, rotated rx 150.39 ry -54.39 rz -78.94 deg; joints [56.788, 29.546, -40.316, -60.768, -77.231, 148.991]
  MoveL 145 to (390.67, 71.76, 229.03) mm, rotated rx 150.39 ry -54.39 rz -78.94 deg; joints [56.632, 29.182, -40.545, -60.725, -77.223, 149.256]
  MoveL 146 to (393.62, 71.59, 229.03) mm, rotated rx 150.39 ry -54.39 rz -78.94 deg; joints [56.491, 28.91, -40.715, -60.678, -77.233, 149.462]
  MoveL 147 to (396.38, 71.57, 229.03) mm, rotated rx 150.39 ry -54.39 rz -78.94 deg; joints [56.348, 28.664, -40.868, -60.627, -77.252, 149.652]
  MoveL 148 to (398.78, 71.57, 229.03) mm, rotated rx 150.39 ry -54.39 rz -78.94 deg; joints [56.221, 28.453, -40.999, -60.58, -77.272, 149.818]
  MoveL 149 to (401.85, 71.57, 229.03) mm, rotated rx 150.39 ry -54.39 rz -78.94 deg; joints [56.057, 28.182, -41.165, -60.519, -77.298, 150.028]
  MoveL 150 to (405.71, 71.57, 229.03) mm, rotated rx 150.39 ry -54.39 rz -78.94 deg; joints [55.849, 27.844, -41.371, -60.439, -77.332, 150.291]
  MoveL 151 to (409.94, 71.57, 229.03) mm, rotated rx 150.39 ry -54.39 rz -78.94 deg; joints [55.619, 27.475, -41.595, -60.35, -77.372, 150.578]
  Establecer velocidad (1000.0 mm/s)
  MoveL 152 to (409.94, 71.57, 229.03) mm, rotated rx 150.39 ry -54.39 rz -78.94 deg; joints [55.619, 27.475, -41.595, -60.35, -77.372, 150.578]
  MoveL 153 to (429.55, 71.57, 327.09) mm, rotated rx 150.39 ry -54.39 rz -78.94 deg; joints [54.514, 19.004, -30.081, -58.15, -84.045, 141.022]

